(* IEC 61131-3 sources: daoli-st-library/DL_Device (part 34) *)

(* ---- FB_DL_VacuumEjector.st ---- *)
(*==============================================================================
 * 组件名称 (Component)  : FB_DL_VacuumEjector
 * 所属子库 (Sublibrary) : DL_Device
 * 当前版本 (Version)    : 1.0.1
 * 兼容性   (Platform)   : CODESYS 3.5 / TwinCAT 3 / 汇川 InoProShop / Machine Expert
 *                         仅依赖 Standard.library（TON / R_TRIG / TP），零厂商方言
 * 分类     (Category)   : 设备执行器功能块（Function Block，实现 I_DL_VacuumGenerator）
 * 功能简述 (Function)   : 真空发生器（射流式负压源）控制功能块。负压阈值
 *                         建立判据（负压域迟滞：建立用设定值、保持放宽
 *                         迟滞带防临界抖动）+ 可选真空开关双确认；破真空
 *                         吹气定宽单发脉冲（吹气期间真空阀强制断）；负压
 *                         反馈非有限值防御保持末次有效值；建立超时锁存；
 *                         状态机 ENUM + CASE + ELSE 兜底。
 * 接口实现 (Implements) : I_DL_VacuumGenerator。接口 OUT 列同名成员
 *                         （eState/bVacuumOk/fPressure/bFault/uErrorId）按
 *                         R22 以只读 PROPERTY GET 承载（内部镜像同源），
 *                         非接口成员 bVacuumValve/bBlowValve/bHolding 保留
 *                         VAR_OUTPUT；方法 CmdEvacuate/CmdBlowOff/CmdStop/
 *                         CmdReset 全部在本文件尾部落地。
 * 开源溯源 (Origin)     : 来源标签 lbp-device（RAW_NOTES_R6 S-1：真空吸持的
 *                         建立-保持迟滞判据、破真空吹气定宽脉冲、真空开关
 *                         双确认等行业公知工程惯例，公开教学资料，仅借鉴
 *                         通用工程语义；状态机、迟滞方向、故障码按本库红线
 *                         独立设计，clean-room 未复制源码）。
 * 红线自检 (Redline)    : R1 零全局变量表/外部变量引用 ✓｜R2 零物理 IO 地址 ✓
 *                         R3 纯 IEC 61131-3 ✓｜R4 防除零/非有限值防御/浮点
 *                         容差比较 ✓｜R5 全变量中英双语同行注释 ✓
 *                         R6 ENUM+CASE+ELSE ✓｜R7 六个定时器/边缘/脉冲实例
 *                         主体最前部无条件刷新 ✓
 * 公约遵循 (Convention) : 0.1/R23 本块为事件型状态机 + 逐拍组合阈值判定：
 *                         迟滞保持态每拍由实时负压重算自校正，无积分/滤波
 *                         类需要首扫初始化的连续量驻留状态，免首扫（无
 *                         bInit 标志）。
 *                         0.7 故障码段位 16#0003_xxxx：【故障级】0003_0230
 *                         负压反馈信号无效 / 0003_0231 真空建立超时（含
 *                         双确认模式下开关校验超窗）/ 0003_0232 非法状态，
 *                         全部 R15 锁存仅复位可清；本块无信息级码，bFault
 *                         派生式天然排除信息级（0.2）。
 * 偏离留档 (Deviation)  : 依 R11 头注释留档，共 1 条：
 *                         ① 规格建议吹气脉冲用"内部时间戳累积法"自实现
 *                           TP 语义；时间戳累积需时钟基准，与公约 0.9
 *                           "禁读时钟、时间一律注入"冲突，本实现改用
 *                           IEC 标准 TP 定宽脉冲定时器（Standard.library，
 *                           纯跨平台，语义等价），R14 断输入一拍规则对
 *                           组态期定值 PT 不涉及。
 * 修订历史 (Revision)   :
 *   2026-11-15  v1.0.0  首版入库（R6 轮 · DL_Device 阀门/驱动族深化）
 *   2026-11-15  v1.0.1  终审修复【致命】吹气脉冲触发时序：原实现 _bBlowReq
 *                       于主体末尾同拍自清，TP 实例（段 1 最前部刷新）永远
 *                       采不到 TRUE 入参，bBlowValve 恒 FALSE、eBlowing 态
 *                       下一拍即退回 eIdle（验收向量 V3 不成立，R13 逐拍
 *                       推演复现）。修法：自清动作移至 TP 实例调用之后，
 *                       TP 本拍采样 TRUE 起振、下一拍入参回落，定宽脉冲
 *                       由 TP 自身保持。引脚契约零变更。
 *============================================================================*)
FUNCTION_BLOCK FB_DL_VacuumEjector IMPLEMENTS I_DL_VacuumGenerator
VAR_INPUT
    bCmdEvacuate      : BOOL;           // 建立真空指令（Evacuate command），上升沿生效 / Evacuate command, rising edge effective
    bCmdBlowOff       : BOOL;           // 破真空吹气指令（Blow-off command），上升沿生效，输出 tBlowPulse 定宽脉冲 / Blow-off command, rising edge outputs fixed-width pulse
    fPressureFeedback : REAL;           // 负压表反馈（Pressure feedback）[kPa]，0=大气，负值=真空度；非有限值防御 / Pressure feedback [kPa], 0 = atmospheric, negative = vacuum, non-finite defended
    bFbVacuumSwitch   : BOOL;           // 可选真空开关反馈（Optional vacuum switch feedback），TRUE=真空确认 / Optional vacuum switch feedback, TRUE = vacuum confirmed
    bUseSensorCheck   : BOOL;           // 开关反馈校验使能（Sensor check enable），TRUE=负压阈值+开关双确认 / Sensor check enable, TRUE = threshold + switch dual confirmation
    fVacuumSetpoint   : REAL := -60.0;  // 真空建立阈值（Vacuum setpoint）[kPa]，负压域 / Vacuum establishment threshold in negative-pressure domain
    fVacuumHysteresis : REAL := 5.0;    // 真空判定迟滞（Vacuum hysteresis）[kPa]，保持判据放宽量，负值防御钳零 / Hysteresis band for hold criterion, negative clamped to zero
    tEstablishTimeout : TIME := T#5S;   // 真空建立超时（Establish timeout），T#0S=禁用 / Establish timeout, T#0S disables the check
    tBlowPulse        : TIME := T#500MS; // 破真空吹气脉冲宽度（Blow-off pulse width）/ Blow-off pulse width
    tDebounce         : TIME := T#20MS; // 开关反馈防抖（Switch debounce），T#0S=直通 / Switch feedback debounce, T#0S = pass-through
    bReset            : BOOL;           // 故障复位（Fault reset），上升沿生效 / Fault reset, rising edge effective
END_VAR

VAR_OUTPUT
    bVacuumValve : BOOL;                // 真空电磁阀输出（Vacuum solenoid valve），TRUE=抽真空 / Vacuum solenoid valve, TRUE = evacuating
    bBlowValve   : BOOL;                // 破真空吹气阀输出（Blow-off solenoid valve），定宽脉冲 / Blow-off solenoid valve, fixed-width pulse
    bHolding     : BOOL;                // 吸附保持中指示（Holding indicator），真空确认态为 TRUE / Holding indicator, TRUE in vacuum-ok state
END_VAR

VAR
    _eState         : E_DL_VacuumState := E_DL_VacuumState.eIdle; // 内部状态机步序（Internal state step），外部经属性只读 / Internal state, read-only via property
    _bFaultLatch    : BOOL;           // 故障锁存标志（Fault latch flag），仅复位清除 / Fault latch flag, cleared only by reset
    _uErrorIdInt    : UDINT;          // 内部故障码寄存（Internal error register），随锁存写入 / Internal error register written on latch
    _bPendEvac      : BOOL;           // 方法抽真空请求（Method evacuate request），由 CmdEvacuate 置位 / Method evacuate request set by CmdEvacuate
    _bPendBlow      : BOOL;           // 方法吹气请求（Method blow-off request），由 CmdBlowOff 置位 / Method blow-off request set by CmdBlowOff
    _bPendStop      : BOOL;           // 方法停止请求（Method stop request），由 CmdStop 置位 / Method stop request set by CmdStop
    _bPendReset     : BOOL;           // 方法复位请求（Method reset request），由 CmdReset 置位 / Method reset request set by CmdReset
    _bBlowReq       : BOOL;           // 吹气单拍触发请求（Blow pulse trigger request），上升沿消费置位一拍 / One-cycle blow trigger, set on edge consumption
    _fPressValid    : REAL := 0.0;    // 末次有效负压值（Last valid pressure）[kPa]，非有限值防御保持载体 / Last valid pressure hold carrier
    _fSetpEff       : REAL := -60.0;  // 防御后建立阈值（Sanitized setpoint）[kPa] / Sanitized vacuum setpoint
    _fHystEff       : REAL := 5.0;    // 防御后迟滞带（Sanitized hysteresis）[kPa]，钳制非负 / Sanitized hysteresis band, clamped non-negative
    _bPressValid    : BOOL;           // 本拍负压输入有效性（Pressure input validity this cycle），非有限值为 FALSE / FALSE when pressure input non-finite
    _bSwFilt        : BOOL;           // 防抖后真空开关（Debounced vacuum switch）/ Debounced vacuum switch signal
    _bInEstablish   : BOOL;           // 建立超时计时条件（Establish timeout timing condition）/ Timing condition of establish timeout
    _bEstToEn       : BOOL;           // 建立超时使能（Establish timeout enable），参数大于零有效 / Establish timeout enable, active when above zero
    _bEstablished   : BOOL;           // 本拍真空建立判据结果（Establishment criterion result this cycle）/ Establishment criterion result this cycle
    _bHoldCriterion : BOOL;           // 本拍保持判据结果（Hold criterion result this cycle），迟滞放宽域 / Hold criterion result within hysteresis band
    _fbTrigEvac     : R_TRIG;         // 引脚抽真空指令上升沿（Pin evacuate command edge）/ Pin evacuate command rising edge
    _fbTrigBlow     : R_TRIG;         // 引脚吹气指令上升沿（Pin blow-off command edge）/ Pin blow-off command rising edge
    _fbTrigReset    : R_TRIG;         // 引脚复位上升沿（Pin reset edge）/ Pin reset rising edge
    _fbTonSwDeb     : TON;            // 真空开关防抖定时器（Vacuum switch debounce timer）/ Vacuum switch debounce timer instance
    _fbTonEstablish : TON;            // 真空建立超时定时器（Establish timeout timer）/ Establish timeout timer instance
    _fbTpBlow       : TP;             // 吹气定宽脉冲定时器（Blow-off pulse timer），IEC 标准 TP / Blow-off fixed-width pulse timer, IEC standard TP
END_VAR

METHOD CmdEvacuate : BOOL
VAR_INPUT
END_VAR
IF _bFaultLatch OR (_eState = E_DL_VacuumState.eFault) THEN
    CmdEvacuate := FALSE;     // 故障态拒绝（Rejected in fault state）
ELSE
    _bPendEvac  := TRUE;      // 登记抽真空请求，主体状态机消化（Register evacuate request, consumed by body）
    CmdEvacuate := TRUE;      // 受理成功（Accepted）
END_IF

(*------------------------------------------------------------------------------
 * 方法: CmdBlowOff —— 破真空吹气指令（单发定宽脉冲）。故障态拒绝。
 *      Method CmdBlowOff - blow-off command (one-shot pulse), rejected in fault.
 *------------------------------------------------------------------------------*)
    END_METHOD

METHOD CmdBlowOff : BOOL
VAR_INPUT
END_VAR
IF _bFaultLatch OR (_eState = E_DL_VacuumState.eFault) THEN
    CmdBlowOff := FALSE;      // 故障态拒绝（Rejected in fault state）
ELSE
    _bPendBlow := TRUE;       // 登记吹气请求，主体状态机消化（Register blow request, consumed by body）
    CmdBlowOff := TRUE;       // 受理成功（Accepted）
END_IF

(*------------------------------------------------------------------------------
 * 方法: CmdStop —— 双阀全断保持现状。故障态拒绝返回 FALSE。
 *      Method CmdStop - both valves off and hold, rejected with FALSE in fault.
 *------------------------------------------------------------------------------*)
    END_METHOD

METHOD CmdStop : BOOL
VAR_INPUT
END_VAR
IF _bFaultLatch OR (_eState = E_DL_VacuumState.eFault) THEN
    CmdStop := FALSE;         // 故障态拒绝（Rejected in fault state）
ELSE
    _bPendEvac := FALSE;      // 注销全部动作请求（Cancel all action requests）
    _bPendBlow := FALSE;
    _bPendStop := TRUE;       // 登记停止请求，主体状态机消化（Register stop request, consumed by body）
    CmdStop    := TRUE;       // 受理成功（Accepted）
END_IF

(*------------------------------------------------------------------------------
 * 方法: CmdReset —— 复位故障，返回是否可复位（存在锁存故障时为 TRUE）。
 *      Method CmdReset - reset fault, returns TRUE only when a latch exists.
 *------------------------------------------------------------------------------*)
    END_METHOD

METHOD CmdReset : BOOL
VAR_INPUT
END_VAR
IF _bFaultLatch OR (_eState = E_DL_VacuumState.eFault) THEN
    _bPendReset := TRUE;      // 登记复位请求，主体状态机消化（Register reset request, consumed by body）
    CmdReset    := TRUE;      // 可复位（Resettable）
ELSE
    CmdReset    := FALSE;     // 无故障可复位（Nothing to reset）
END_IF

(*------------------------------------------------------------------------------
 * 属性: eState（GET）—— 当前状态机状态只读视图。
 *      Property eState (GET) - read-only view of the current state machine state.
 *------------------------------------------------------------------------------*)
    END_METHOD

// ============================================================================
// 段 1｜定时器与边缘检测实例无条件周期刷新（R7：严禁置于 IF/CASE 分支内）
//      Unconditional per-cycle refresh of all timer and edge instances (R7)
// ============================================================================
_fbTrigEvac(CLK := bCmdEvacuate);
_fbTrigBlow(CLK := bCmdBlowOff);
_fbTrigReset(CLK := bReset);
_fbTonSwDeb(IN := bFbVacuumSwitch, PT := tDebounce); // 开关持续为真 tDebounce 才确认（Switch must hold TRUE for tDebounce）
_bSwFilt := _fbTonSwDeb.Q;            // 防抖后开关（Debounced switch）
_bEstToEn := (tEstablishTimeout > T#0S); // 超时参数为零 = 自检禁用（Zero timeout = check disabled）
_bInEstablish := (_eState = E_DL_VacuumState.eEvacuating) AND _bEstToEn; // 建立超时计时条件（Timeout timing condition）
_fbTonEstablish(IN := _bInEstablish, PT := tEstablishTimeout);
_fbTpBlow(IN := _bBlowReq, PT := tBlowPulse); // 吹气定宽脉冲（Fixed-width blow pulse, TP semantics）
_bBlowReq := FALSE;                   // 单拍触发请求在 TP 采样后立即自清：TP 于本拍见到
                                      // TRUE 并起振，下一拍入参回落 FALSE，TP 定宽保持
                                      // （One-cycle trigger cleared right after TP sampling,
                                      // pulse held by TP for the full width）

// ============================================================================
// 段 2｜参数防御（0.8：非数自比检测，默认值先赋）+ 迟滞钳零
//      Parameter sanitation (0.8 NaN self-compare, defaults first) + clamp
// ============================================================================
_fSetpEff := fVacuumSetpoint;         // 建立阈值镜像（Setpoint mirror）
IF _fSetpEff <> _fSetpEff THEN        // 非数自比检测（NaN self-compare test）
    _fSetpEff := -60.0;               // 回落默认阈值（Fallback to default setpoint）
END_IF
_fHystEff := fVacuumHysteresis;       // 迟滞带镜像（Hysteresis mirror）
IF _fHystEff <> _fHystEff THEN        // 非数自比检测（NaN self-compare test）
    _fHystEff := 5.0;                 // 回落默认迟滞（Fallback to default hysteresis）
END_IF
IF _fHystEff < 0.0 THEN
    _fHystEff := 0.0;                 // 负迟滞会收窄判定域，钳零防错（Negative band narrows domain, clamp to zero）
END_IF

// ============================================================================
// 段 3｜负压输入有效性全局监视（优先级最高，吸附安全相关故为故障级）
//      Pressure validity global monitor (highest priority, fault level due
//      to holding safety relevance)
// ============================================================================
_bPressValid := (fPressureFeedback = fPressureFeedback); // 非数自比检测：等号成立即有效（NaN iff self-compare fails）
IF _bPressValid THEN
    _fPressValid := fPressureFeedback; // 更新末次有效负压（Update last valid pressure）
ELSE
    _bFaultLatch := TRUE;              // 反馈失效锁存（Feedback loss latch）
    _uErrorIdInt := 16#0003_0230;      // 0003_0230 负压反馈信号无效【故障级】/ Pressure feedback invalid, fault level
    _eState      := E_DL_VacuumState.eFault; // 强制故障态（Force fault state）
END_IF

// 真空判据（clean-room 内联迟滞语义，负压域方向：值越负真空越强）
// Vacuum criteria (inline hysteresis, negative-pressure domain: more negative = stronger)
_bEstablished := (_fPressValid <= _fSetpEff);                          // 建立判据：达到设定真空（Establish: reached setpoint vacuum）
_bHoldCriterion := (_fPressValid <= (_fSetpEff + _fHystEff));          // 保持判据：迟滞带放宽防临界抖动（Hold: widened by hysteresis band）

// ============================================================================
// 段 4｜核心状态机（ENUM + CASE，含 ELSE 非法状态兜底）
//      Core state machine (ENUM + CASE with ELSE illegal-state fallback)
// ============================================================================
IF _bFaultLatch OR (_eState = E_DL_VacuumState.eFault) THEN
    // 故障锁存态：清空全部请求，仅复位可退出（Latched fault: requests cleared, reset-only exit）
    _bPendEvac  := FALSE;             // 清方法请求（Clear method requests）
    _bPendBlow  := FALSE;
    _bPendStop  := FALSE;
    _bBlowReq   := FALSE;             // 撤销未触发脉冲请求（Cancel pending pulse trigger）
    IF _bPendReset OR _fbTrigReset.Q THEN
        _bPendReset  := FALSE;        // 消费复位请求（Consume reset request）
        _bFaultLatch := FALSE;        // 解除锁存（Release latch）
        _uErrorIdInt := 0;            // 故障码清零（Error code cleared）
        _eState      := E_DL_VacuumState.eIdle; // 回空闲态（Back to idle）
    END_IF
ELSE
    IF _bPendReset OR _fbTrigReset.Q THEN
        _bPendReset := FALSE;         // 无故障时消化复位请求（Absorb reset request when no fault）
    END_IF
    CASE _eState OF

        E_DL_VacuumState.eIdle: // 空闲稳态：双阀全断
            IF _bPendEvac OR _fbTrigEvac.Q THEN
                _bPendEvac := FALSE;            // 消费抽真空请求（Consume evacuate request）
                _eState    := E_DL_VacuumState.eEvacuating; // 转抽真空（To evacuating）
            ELSIF _bPendBlow OR _fbTrigBlow.Q THEN
                _bPendBlow := FALSE;            // 消费吹气请求（Consume blow request）
                _bBlowReq  := TRUE;             // 触发定宽脉冲（Trigger fixed-width pulse）
                _eState    := E_DL_VacuumState.eBlowing;
            ELSIF _bPendStop THEN
                _bPendStop := FALSE;            // 空闲态消化停止请求（Absorb stop request in idle）
            END_IF

        E_DL_VacuumState.eEvacuating: // 抽真空中：真空阀开，等待建立确认
            IF _bPendBlow OR _fbTrigBlow.Q THEN
                _bPendBlow := FALSE;            // 中途改吹气（Mid-way blow-off）
                _bBlowReq  := TRUE;
                _eState    := E_DL_VacuumState.eBlowing;
            ELSIF _bPendStop THEN
                _bPendStop := FALSE;            // 停止：双阀全断（Stop: both valves off）
                _eState    := E_DL_VacuumState.eIdle;
            ELSIF bUseSensorCheck AND _bEstablished AND (NOT _bSwFilt) THEN
                // 阈值达成但开关未确认：继续抽气等待（Threshold reached, switch pending: keep evacuating）
            ELSIF (NOT bUseSensorCheck) AND _bEstablished THEN
                _eState := E_DL_VacuumState.eVacuumOk; // 纯阈值模式：建立确认（Pure threshold: established）
            ELSIF bUseSensorCheck AND _bEstablished AND _bSwFilt THEN
                _eState := E_DL_VacuumState.eVacuumOk; // 双确认模式：阈值+开关齐备（Dual confirm: threshold AND switch）
            ELSIF _fbTonEstablish.Q THEN
                _bFaultLatch := TRUE;           // 建立超时锁存（Establish timeout latch）
                _uErrorIdInt := 16#0003_0231;   // 0003_0231 真空建立超时/反馈校验失败【故障级】/ Establish timeout or check failure, fault level
                _eState      := E_DL_VacuumState.eFault;
            END_IF

        E_DL_VacuumState.eVacuumOk: // 真空保持态：吸附保持中
            IF _bPendBlow OR _fbTrigBlow.Q THEN
                _bPendBlow := FALSE;            // 破真空放料（Release workpiece by blow-off）
                _bBlowReq  := TRUE;
                _eState    := E_DL_VacuumState.eBlowing;
            ELSIF _bPendStop THEN
                _bPendStop := FALSE;            // 停止：双阀全断（Stop: both valves off）
                _eState    := E_DL_VacuumState.eIdle;
            ELSIF NOT _bHoldCriterion THEN
                _eState := E_DL_VacuumState.eEvacuating; // 真空丢失（超迟滞带）：自动重建（Vacuum lost beyond band: auto re-establish）
            ELSIF bUseSensorCheck AND (NOT _bSwFilt) THEN
                _eState := E_DL_VacuumState.eEvacuating; // 双确认模式下开关脱开：自动重建（Switch dropped in dual mode: re-establish）
            END_IF

        E_DL_VacuumState.eBlowing: // 吹气中：吹气阀定宽脉冲，真空阀强制断
            IF _bPendBlow OR _fbTrigBlow.Q THEN
                _bPendBlow := FALSE;            // 吹气中重复触发忽略（Retrigger ignored while blowing）
            ELSIF _bPendStop THEN
                _bPendStop := FALSE;            // 停止请求提前截断脉冲（Stop request truncates pulse early）
                _bBlowReq  := FALSE;
                _eState    := E_DL_VacuumState.eIdle;
            ELSIF NOT _fbTpBlow.Q THEN
                _eState := E_DL_VacuumState.eIdle; // 脉冲宽度计满自动回空闲（Pulse completed, back to idle）
            END_IF

        ELSE // 非法状态兜底：任何越界枚举值强制锁存故障（Illegal state fallback）
            _bFaultLatch := TRUE;               // 故障锁存（Fault latched）
            _uErrorIdInt := 16#0003_0232;       // 0003_0232 非法状态【故障级】/ Illegal state, fault level
            _eState      := E_DL_VacuumState.eFault;
    END_CASE
END_IF

// ============================================================================
// 段 5｜阀输出推导 + 出口断言（硬约束：吹气期间真空阀必断；故障/空闲双阀必断）
//      Valve output derivation + exit assertions (vacuum valve forced off
//      while blowing; both valves off in fault/idle)
// ============================================================================
bVacuumValve := (_eState = E_DL_VacuumState.eEvacuating) OR (_eState = E_DL_VacuumState.eVacuumOk); // 抽真空与保持期真空阀开（Valve open while evacuating/holding）
bBlowValve := (_eState = E_DL_VacuumState.eBlowing) AND _fbTpBlow.Q; // 吹气阀随 TP 定宽脉冲（Blow valve follows TP pulse）
IF (_eState = E_DL_VacuumState.eBlowing) OR (_eState = E_DL_VacuumState.eFault)
   OR (_eState = E_DL_VacuumState.eIdle) THEN
    bVacuumValve := FALSE;              // 出口断言：吹气/故障/空闲真空阀必断（Assertion: vacuum valve off in blowing/fault/idle）
END_IF

(*------------------------------------------------------------------------------
 * 方法: CmdEvacuate —— 建立真空指令（单发）。故障态一律拒绝返回 FALSE。
 *      Method CmdEvacuate - evacuate command (one-shot), rejected with FALSE in fault.
 *------------------------------------------------------------------------------*)

PROPERTY eState : E_DL_VacuumState
eState := _eState;            // 返回内部状态（Return internal state）

(*------------------------------------------------------------------------------
 * 属性: bVacuumOk（GET）—— 真空建立确认（吸附保持态为 TRUE）。
 *      Property bVacuumOk (GET) - vacuum established (TRUE in holding state).
 *------------------------------------------------------------------------------*)
PROPERTY bVacuumOk : BOOL
bVacuumOk := (_eState = E_DL_VacuumState.eVacuumOk); // 显式状态派生式（Explicit state-derived form）

(*------------------------------------------------------------------------------
 * 属性: fPressure（GET）—— 负压反馈值 [kPa]，0=大气压，负值=真空度。
 *      Property fPressure (GET) - pressure feedback [kPa], 0 = atmospheric, negative = vacuum.
 *------------------------------------------------------------------------------*)
PROPERTY fPressure : REAL
fPressure := _fPressValid;    // 返回末次有效负压保持值（Return last valid pressure hold value）

(*------------------------------------------------------------------------------
 * 属性: bFault（GET）—— 故障锁存指示（信息级码不置本位，0.2 公约）。
 *      Property bFault (GET) - fault latch indicator, info-level codes excluded.
 *------------------------------------------------------------------------------*)
PROPERTY bFault : BOOL
bFault := _bFaultLatch OR (_eState = E_DL_VacuumState.eFault); // 显式排除信息级派生式（Explicit derived form excluding info codes）

(*------------------------------------------------------------------------------
 * 属性: uErrorId（GET）—— 末次故障码（0=无故障）。
 *      Property uErrorId (GET) - last error code (0 = none).
 *------------------------------------------------------------------------------*)
PROPERTY uErrorId : UDINT
uErrorId := _uErrorIdInt;     // 返回内部故障码寄存（Return internal error register）
END_FUNCTION_BLOCK

(* ---- FB_DL_VacuumPumpBasePress.st ---- *)
(*
  Component : FB_DL_VacuumPumpBasePress
  Category  : DL_Device
  Type      : FB
  Version   : 1.0.0
  CodeSeg   : 16#03_1_03
  Summary   : 真空泵本底压强与恢复时间台账：本底压强滑动平均平滑 + 起泵恢复超时事件计数留痕。
              Vacuum pump base pressure and recovery ledger: moving-average smoothing plus restart recovery timeout counting.
  溯源声明  : 道莅自研 clean-room
  边界安全  : 压强非物理域闸（负压 < 0 拦截，非有限 NaN/Inf 拦截）；MA 环形缓冲点数域闸（2..16，防越界）；
              采样窗/恢复窗时长正域闸（> 0）；MA 采样窗与恢复计时窗为独立 TON 实例；
              恢复超时计数用事件触发（timing 停止后不重复累加）；锁存故障有可达清码路径（恢复成功即清）。
  复用      : 无
*)

FUNCTION_BLOCK FB_DL_VacuumPumpBasePress
VAR_INPUT
    bRun       : BOOL;                  (* 监视使能 · Enable *)
    bPumpRun   : BOOL;                  (* 泵运行反馈 [开关]，上升沿起恢复计时 · Pump run feedback *)
    fPressKpa  : LREAL;                 (* 泵入口压强 [kPa] · Pump inlet pressure *)
    fBaseOkKpa : LREAL := 5.0;          (* 本底压强达标阈 [kPa] · Base pressure target *)
    tMaWinMs   : TIME  := T#2000MS;     (* MA 采样节拍 [ms] · MA sample pace *)
    tRecWinMs  : TIME  := T#60000MS;    (* 恢复计时窗 [ms] · Recovery timing window *)
    nMaPts     : INT   := 8;            (* MA 有效点数 [点]，域 2 到 16 · MA valid points *)
    fEps       : LREAL := 1.0E-6;       (* 浮点判零容差 [实数域] · Floating zero tolerance *)
END_VAR
VAR_OUTPUT
    fMaKpa      : LREAL;                (* 本底压强滑动平均 [kPa] · Moving average pressure *)
    bRecTiming  : BOOL;                 (* 恢复计时进行中 [开关] · Recovery timing active *)
    bRecOk      : BOOL;                 (* 最近一次恢复成功 [开关] · Last recovery succeeded *)
    nRecTimeout : UDINT;                (* 恢复超时累计 [次]，事件计数防回卷 · Recovery timeout count *)
    bError      : BOOL;                 (* 故障标志，与故障码配对 · Fault flag paired with codes *)
    uErrorId    : UDINT;                (* 事件码 16#0000_0103，0 无事件 · Event code *)
END_VAR
VAR
    uCode    : WORD;    (* 码位暂存，每拍重算 [码] · Code staging *)
    tonMa    : TON;     (* MA 采样节拍 [ms]，自复位振荡 · MA pace timer, self-reset *)
    tonRec   : TON;     (* 恢复计时窗 [ms]，独立实例 · Recovery window timer, separate instance *)
    rTrigRun : R_TRIG;  (* 起泵上升沿 · Pump start rising edge *)
    aRing    : ARRAY[1..16] OF LREAL;   (* MA 环形缓冲 [kPa] · MA ring buffer *)
    nHead    : INT;     (* 环形头下标 [索引] · Ring head index *)
    nFill    : INT;     (* 已填充点数 [点] · Filled point count *)
    fSum     : LREAL;   (* 环内累加和 [kPa] · Ring sum *)
    bRecFlt  : BOOL;    (* 恢复超时锁存 · Recovery timeout latched *)
    bSigOk   : BOOL;    (* 输入有效标志 · Input validity flag *)
    bTick    : BOOL;    (* 采样到点脉冲 [脉冲] · Sample tick pulse *)
    nI       : INT;     (* 求和循环下标 [索引] · Sum loop index *)
END_VAR
VAR CONSTANT
    DL_VBP_NMAX : INT := 16;            (* 环形缓冲容量 [点] · Ring capacity *)
END_VAR

(* === 段 0 · 实例刷新（每拍无条件，红线 7）=== *)
tonMa(IN := NOT tonMa.Q, PT := tMaWinMs);       (* 采样节拍自复位振荡 / Self-reset MA pace *)
tonRec(IN := bRecTiming, PT := tRecWinMs);      (* 恢复计时窗独立实例 / Separate recovery window *)
rTrigRun(CLK := bPumpRun);                      (* 起泵沿检测 / Pump start edge *)
bTick := tonMa.Q;                               (* 采样脉冲 / Sample tick *)

(* === 段 1 · 输入校验与量程闸 === *)
uCode := 16#0000;                       // 每拍清码（可达清零基线）/ Clear codes each scan
bSigOk := (fPressKpa = fPressKpa) AND (ABS(fPressKpa) < 1.0E308)    // 非有限拦截 / Non-finite guard
          AND (fPressKpa >= 0.0)                                     // 压强非负域闸 / Non-negative pressure
          AND (nMaPts >= 2) AND (nMaPts <= DL_VBP_NMAX)              // 点数域闸，防越界 / Point-count gate
          AND (tMaWinMs > T#0MS) AND (tRecWinMs > T#0MS);            // 窗时长正域闸 / Window duration gates
IF NOT bSigOk THEN
    uCode := 16#0103;                   // 故障级：域外，台账冻结 / Fault: domain invalid
END_IF

(* === 段 2 · 主逻辑：MA 平滑与恢复台账 === *)
IF bSigOk THEN
    IF bTick THEN                       (* 采样到点：写环并重算均值 / Sample tick: write ring *)
        IF nFill < nMaPts THEN
            nFill := nFill + 1;         (* 未满先增填充数 / Grow fill count *)
        ELSE
            fSum := fSum - aRing[nHead];    (* 满环先减旧值 / Remove the old value *)
        END_IF
        aRing[nHead] := fPressKpa;      (* 写入新采样 / Write the new sample *)
        fSum := fSum + fPressKpa;       (* 累加新值 / Add the new value *)
        nHead := (nHead MOD DL_VBP_NMAX) + 1;   (* 头下标循环推进 / Advance the head *)
    END_IF
    IF nFill >= 2 THEN
        fMaKpa := fSum / UDINT_TO_LREAL(INT_TO_UDINT(nFill));   (* 均值，填充数 ≥2 已闸 / Mean *)
    END_IF
    (* 恢复台账：起泵沿起计时，达标即成功，超窗即超时计数 / Recovery ledger *)
    IF rTrigRun.Q THEN
        bRecTiming := TRUE;             (* 拍 N 起泵沿进入，本拍置计时，拍 N+1 tonRec 生效 / Start timing *)
        bRecOk := FALSE;                (* 新恢复未达标 / New recovery pending *)
    END_IF
    IF bRecTiming AND (fMaKpa <= fBaseOkKpa) AND (nFill >= nMaPts) THEN
        bRecTiming := FALSE;            (* 达标：停止计时 / Reached target: stop timing *)
        bRecOk := TRUE;                 (* 恢复成功 / Recovery succeeded *)
        bRecFlt := FALSE;               (* 超时锁存清码（可达路径）/ Reachable clear of the latch *)
    END_IF
    IF bRecTiming AND tonRec.Q THEN     (* 计时窗满仍未达标 / Window expired without target *)
        bRecTiming := FALSE;            (* 停止计时，防重复计数 / Stop timing, no double count *)
        bRecFlt := TRUE;                (* 超时锁存 / Latch the timeout *)
        IF nRecTimeout < 4294967290 THEN
            nRecTimeout := nRecTimeout + 1;     (* 事件计数，一次恢复只计一次 / Count once per recovery *)
        END_IF
    END_IF
END_IF

(* === 段 3 · 输出映射与故障码 === *)
IF NOT bRun THEN
    bRecTiming := FALSE;                (* 撤使能停计时 / Stop timing on disable *)
END_IF
bError := bRecFlt OR (uCode <> 16#0000);        (* 故障标志：超时锁存或域外 / Fault flag *)
IF bRecFlt THEN
    uErrorId := WORD_TO_UDINT(16#0103); (* 码位 16#0000_0103 恢复超时锁存 / Recovery timeout code *)
ELSE
    uErrorId := WORD_TO_UDINT(uCode);   (* 域外码或零 / Domain code or zero *)
END_IF
END_FUNCTION_BLOCK

(* ---- FB_DL_ValveCycleCountBank.st ---- *)
//==============================================================================
// 功能块：FB_DL_ValveCycleCountBank ｜ 中文名称：多阀动作计数寿命台账组
// 所属子库：DL_Device ｜ 版本：v1.0.0 ｜ 日期：2026-11-23
// 兼容：CODESYS V3.5+ / TwinCAT 3 / 汇川 InoProShop（纯标准库 R_TRIG）
// 功能描述：4 阀动作计数寿命台账 Bank：每通道对阀指令上升沿计数（全行程
//           动作次数），独立维护阈值（UDINT），计数达阈值置该通道维护预警
//           bMaintX（不置故障——维护预警是台账事实非软件错误）。计数饱和
//           于 UDINT 上限 4294967295 不回绕（信息级留痕），复位经 bRst 沿
//           或 bRstChX 单通道沿。
//           同族分工：单阀寿命判定（阀位双阈值跨越 + 双源同证去抖 + 分级
//           预警）属 FB_DL_ValveCycleLifeCounter；本件为 4 通道指令沿计数
//           Bank 台账（无反馈口径），互不替代（R73 互引）。
// 开源溯源 (Origin)：原创实现（t2-2-lbp 阀诊断深化，零外部源码行，clean-room
//           独立编写）
// 公开接口清单：输入 {bCmdCh1..4, uLimitCh1..4} / bRst / bRstCh1..4；
//               输出 {uCntCh1..4, bMaintCh1..4} / uErrCode / bValid
// 错误码表：16#0003_0754 信息级（任一通道计数饱和不回绕，不置 bError）/
//           16#0003_0755 预留禁用（不得挪用）
// 状态机：N/A（台账计数无状态机；R_TRIG ×8 每拍无条件刷新）
// 边界行为：① 计数饱和于 4294967295 不回绕（信息级 0754 留痕）；
//           ② R_TRIG 全部每拍无条件刷新（不入分支，红线 R7）；
//           ③ 维护预警随计数回落自动撤销（阈值比较瞬时量，不锁存）；
//           ④ 复位沿仅清计数，不清阈值与信息码（信息码每拍重算）。
// 修订历史：v1.0.0 2026-11-23 首版（R73 派单 · 批 3 · 序 16）
//==============================================================================

(*==============================================================================
 * 功能块: FB_DL_ValveCycleCountBank
 * 调用约定: 每个扫描周期无条件调用一次；实例状态全部驻留于私有变量。
 *==============================================================================*)
FUNCTION_BLOCK FB_DL_ValveCycleCountBank
VAR_INPUT
    bCmdCh1  : BOOL := FALSE;          // 阀 1 指令（上升沿 = 一次全行程动作）/ Valve 1 command, rising edge = one full stroke
    bCmdCh2  : BOOL := FALSE;          // 阀 2 指令（上升沿计数）/ Valve 2 command, counted on rising edge
    bCmdCh3  : BOOL := FALSE;          // 阀 3 指令（上升沿计数）/ Valve 3 command, counted on rising edge
    bCmdCh4  : BOOL := FALSE;          // 阀 4 指令（上升沿计数）/ Valve 4 command, counted on rising edge
    uLimitCh1: UDINT := 1000000;       // 阀 1 维护阈值 [次] / Valve 1 maintenance threshold [cycles]
    uLimitCh2: UDINT := 1000000;       // 阀 2 维护阈值 [次] / Valve 2 maintenance threshold [cycles]
    uLimitCh3: UDINT := 1000000;       // 阀 3 维护阈值 [次] / Valve 3 maintenance threshold [cycles]
    uLimitCh4: UDINT := 1000000;       // 阀 4 维护阈值 [次] / Valve 4 maintenance threshold [cycles]
    bRst     : BOOL := FALSE;          // 全组复位（上升沿，清全部计数）/ Bank reset, rising edge, clears all counts
    bRstCh1  : BOOL := FALSE;          // 阀 1 单通道复位沿 / Valve 1 channel reset edge
    bRstCh2  : BOOL := FALSE;          // 阀 2 单通道复位沿 / Valve 2 channel reset edge
    bRstCh3  : BOOL := FALSE;          // 阀 3 单通道复位沿 / Valve 3 channel reset edge
    bRstCh4  : BOOL := FALSE;          // 阀 4 单通道复位沿 / Valve 4 channel reset edge
END_VAR
VAR_OUTPUT
    uCntCh1  : UDINT;                  // 阀 1 累计动作数 [次] / Valve 1 accumulated cycles
    uCntCh2  : UDINT;                  // 阀 2 累计动作数 [次] / Valve 2 accumulated cycles
    uCntCh3  : UDINT;                  // 阀 3 累计动作数 [次] / Valve 3 accumulated cycles
    uCntCh4  : UDINT;                  // 阀 4 累计动作数 [次] / Valve 4 accumulated cycles
    bMaintCh1: BOOL;                   // 阀 1 维护预警（计数达阈值）/ Valve 1 maintenance warning
    bMaintCh2: BOOL;                   // 阀 2 维护预警（计数达阈值）/ Valve 2 maintenance warning
    bMaintCh3: BOOL;                   // 阀 3 维护预警（计数达阈值）/ Valve 3 maintenance warning
    bMaintCh4: BOOL;                   // 阀 4 维护预警（计数达阈值）/ Valve 4 maintenance warning
    uErrCode : UDINT;                  // 信息级码，0 = 无信息 / Info-level code, 0 = none
    bValid   : BOOL;                   // 输出可用标志 / Outputs usable flag
END_VAR
VAR
    trigCmd1 : R_TRIG;                 // 阀 1 指令沿检测，每拍无条件刷新 / Valve 1 command edge, refreshed every scan
    trigCmd2 : R_TRIG;                 // 阀 2 指令沿检测，每拍无条件刷新 / Valve 2 command edge, refreshed every scan
    trigCmd3 : R_TRIG;                 // 阀 3 指令沿检测，每拍无条件刷新 / Valve 3 command edge, refreshed every scan
    trigCmd4 : R_TRIG;                 // 阀 4 指令沿检测，每拍无条件刷新 / Valve 4 command edge, refreshed every scan
    trigRst  : R_TRIG;                 // 全组复位沿检测，每拍无条件刷新 / Bank reset edge, refreshed every scan
    trigRst1 : R_TRIG;                 // 阀 1 复位沿检测，每拍无条件刷新 / Valve 1 reset edge, refreshed every scan
    trigRst2 : R_TRIG;                 // 阀 2 复位沿检测，每拍无条件刷新 / Valve 2 reset edge, refreshed every scan
    trigRst3 : R_TRIG;                 // 阀 3 复位沿检测，每拍无条件刷新 / Valve 3 reset edge, refreshed every scan
    trigRst4 : R_TRIG;                 // 阀 4 复位沿检测，每拍无条件刷新 / Valve 4 reset edge, refreshed every scan
END_VAR
VAR CONSTANT
    DL_VCC_MAX     : UDINT := 4294967295; // UDINT 计数上限（饱和不回绕）/ UDINT count ceiling, saturating
    DL_VCC_CODE_SAT: UDINT := 16#0003_0754; // 信息级：计数饱和码 / Info code: count saturated
END_VAR

// ---- 段 1｜沿实例无条件刷新（红线 R7：全部 8 实例不入分支）----
trigCmd1(CLK := bCmdCh1);             // 阀 1 指令沿每拍刷新 / Valve 1 edge refreshed
trigCmd2(CLK := bCmdCh2);             // 阀 2 指令沿每拍刷新 / Valve 2 edge refreshed
trigCmd3(CLK := bCmdCh3);             // 阀 3 指令沿每拍刷新 / Valve 3 edge refreshed
trigCmd4(CLK := bCmdCh4);             // 阀 4 指令沿每拍刷新 / Valve 4 edge refreshed
trigRst(CLK := bRst);                 // 全组复位沿每拍刷新 / Bank reset edge refreshed
trigRst1(CLK := bRstCh1);             // 阀 1 复位沿每拍刷新 / Valve 1 reset edge refreshed
trigRst2(CLK := bRstCh2);             // 阀 2 复位沿每拍刷新 / Valve 2 reset edge refreshed
trigRst3(CLK := bRstCh3);             // 阀 3 复位沿每拍刷新 / Valve 3 reset edge refreshed
trigRst4(CLK := bRstCh4);             // 阀 4 复位沿每拍刷新 / Valve 4 reset edge refreshed

// ---- 段 2｜计数推进：饱和不回绕（信息级留痕，每拍重算）----
IF trigCmd1.Q AND (uCntCh1 < DL_VCC_MAX) THEN
    uCntCh1 := uCntCh1 + 1;           // 阀 1 计数推进 / Valve 1 count advance
END_IF
IF trigCmd2.Q AND (uCntCh2 < DL_VCC_MAX) THEN
    uCntCh2 := uCntCh2 + 1;           // 阀 2 计数推进 / Valve 2 count advance
END_IF
IF trigCmd3.Q AND (uCntCh3 < DL_VCC_MAX) THEN
    uCntCh3 := uCntCh3 + 1;           // 阀 3 计数推进 / Valve 3 count advance
END_IF
IF trigCmd4.Q AND (uCntCh4 < DL_VCC_MAX) THEN
    uCntCh4 := uCntCh4 + 1;           // 阀 4 计数推进 / Valve 4 count advance
END_IF
IF (uCntCh1 = DL_VCC_MAX) OR (uCntCh2 = DL_VCC_MAX)
   OR (uCntCh3 = DL_VCC_MAX) OR (uCntCh4 = DL_VCC_MAX) THEN
    uErrCode := DL_VCC_CODE_SAT;      // 信息级：计数饱和不回绕留痕 / Info: saturation trace, no wrap
END_IF

// ---- 段 3｜复位路径：全组沿 + 单通道沿（锁存声明的清除沿）----
IF trigRst.Q THEN                     // 全组复位沿
    uCntCh1 := 0;                     // 阀 1 计数清零 / Valve 1 count cleared
    uCntCh2 := 0;                     // 阀 2 计数清零 / Valve 2 count cleared
    uCntCh3 := 0;                     // 阀 3 计数清零 / Valve 3 count cleared
    uCntCh4 := 0;                     // 阀 4 计数清零 / Valve 4 count cleared
END_IF
IF trigRst1.Q THEN
    uCntCh1 := 0;                     // 阀 1 单通道清零 / Valve 1 channel clear
END_IF
IF trigRst2.Q THEN
    uCntCh2 := 0;                     // 阀 2 单通道清零 / Valve 2 channel clear
END_IF
IF trigRst3.Q THEN
    uCntCh3 := 0;                     // 阀 3 单通道清零 / Valve 3 channel clear
END_IF
IF trigRst4.Q THEN
    uCntCh4 := 0;                     // 阀 4 单通道清零 / Valve 4 channel clear
END_IF

// ---- 段 4｜维护预警装配：阈值比较瞬时量（随计数回落自动撤销，不锁存）----
bMaintCh1 := uCntCh1 >= uLimitCh1;    // 阀 1 维护预警 / Valve 1 maintenance warning
bMaintCh2 := uCntCh2 >= uLimitCh2;    // 阀 2 维护预警 / Valve 2 maintenance warning
bMaintCh3 := uCntCh3 >= uLimitCh3;    // 阀 3 维护预警 / Valve 3 maintenance warning
bMaintCh4 := uCntCh4 >= uLimitCh4;    // 阀 4 维护预警 / Valve 4 maintenance warning
bValid := TRUE;                       // 台账输出恒可用 / Ledger outputs always usable
END_FUNCTION_BLOCK

(* ---- FB_DL_ValveCycleLifeCounter.st ---- *)
(*
  Name        : FB_DL_ValveCycleLifeCounter
  Category    : DL_Device
  Version     : 1.0.0
  Purpose     : 阀门动作循环寿命计数：行程到位 + 扭角峰值双源同证并经去抖确认才计一个循环，累计数达保养阈值即预警；/ Valve cycle-life counter: one cycle is counted only when both stroke-limit and torque sources agree and the agreement is debounce-confirmed; a maintenance warning is raised at the threshold
  溯源        : 借 t2-8-isa182·回路一致性 的分类/参数域组织，clean-room 实现
  Boundary    : ① 组态闸：保养阈值 < 1 / 去抖时间 <= 0 → 锁存故障（阈值 0 会使预警无意义）；
                ② 双源判据：行程与扭角须同拍同真（AND），单源漂移不会虚计（去抖再拦短时毛刺）；
                ③ 计数用净额单点写入 + 饱和上限（R28 防回绕），不使用 CTU 双向端；
                ④ 循环脉冲 _bCycC 内部置位 → 段 5 统一出口映射单拍（R187），CASE 内不直写出口；
                ⑤ 本件仅计数与预警，不执行保养联锁（属主边界）。
*)
TYPE E_DL_VclState :
(
    eIdle  := 0,                             (* 未使能 / Disabled *)
    eCount := 10,                            (* 寿命计数运行 / Counting *)
    eFault := 90                             (* 故障锁存相 / Fault latched *)
);
END_TYPE

TYPE E_DL_VclCause :
(
    eNone       := 0,                        (* 无故障成因 / No cause *)
    eCfgIllegal := 1,                        (* 组态非法：阈值/去抖越域 / Illegal config *)
    ePhaseBad   := 2                         (* 非法相位兜底 / Illegal phase fallback *)
);
END_TYPE

FUNCTION_BLOCK FB_DL_ValveCycleLifeCounter
VAR_INPUT
    bStrokeOk   : BOOL := FALSE;             (* 行程到位信号（限位开关/位控回读）[-] / Stroke limit reached *)
    bTorqueOk   : BOOL := FALSE;             (* 扭角峰值信号（扭矩/扭角判据回读）[-] / Torque-angle criterion met *)
    tDebounce   : TIME := T#200MS;           (* 双源同证去抖时长，域 > T#0S [ms] / Dual-source debounce time, > 0 *)
    nMaintLimit : UDINT := 100000;           (* 保养阈值（累计循环数），域 >= 1 [次] / Maintenance cycle threshold, >= 1 *)
    bEnable     : BOOL := TRUE;              (* 计数使能 [-] / Enable *)
    bReset      : BOOL := FALSE;             (* 复位命令，上升沿清计数与故障（保养完成侧清零亦可用）[-] / Reset command *)
END_VAR
VAR_OUTPUT
    nCycles     : UDINT;                     (* 累计动作循环数（净额，饱和）[次] / Accumulated cycles, saturated *)
    fCycPct     : REAL;                      (* 寿命消耗百分比 = 计数/阈值（饱和 0..100）[%] / Life consumed percentage *)
    bCycPulse   : BOOL;                      (* 本拍新增一个循环（单拍脉冲）[-] / One new cycle this scan *)
    bMaintWarn  : BOOL;                      (* 保养预警：累计数 >= 阈值（电平，复位沿清）[-] / Maintenance warning level *)
    eState      : E_DL_VclState;             (* 状态出口 / State outlet *)
    eCause      : E_DL_VclCause;             (* 故障成因出口（R190 归因唯一） / Fault cause outlet *)
    bError      : BOOL;                      (* 故障锁存标志 [-] / Fault latch flag *)
END_VAR
VAR
    _eState   : E_DL_VclState := E_DL_VclState.eIdle;    (* 内部相位（CASE 唯一写入目标） / Internal phase *)
    _eCause   : E_DL_VclCause := E_DL_VclCause.eNone;    (* 故障成因锁存量 / Latched cause *)
    rtReset   : R_TRIG;                      (* 复位沿实例，段 0 无条件调用 / Reset edge instance *)
    rtCyc     : R_TRIG;                      (* 去抖确认输出沿实例，段 0 无条件调用 / Debounced-cycle edge *)
    tonDeb    : TON;                         (* 双源同证去抖计时器（IN 由双源派生） / Dual-source debounce timer *)
    _bFault   : BOOL;                        (* 故障锁存位 / Latched fault bit *)
    _bCfgBad  : BOOL;                        (* 组态非法当拍量 / Illegal config this scan *)
    _bDual    : BOOL;                        (* 双源同证当拍量（行程 AND 扭角） / Dual-source agreement this scan *)
    _bCycC    : BOOL;                        (* 循环确认内部单拍量（出口统一映射，R187） / Cycle-confirmed internal pulse *)
END_VAR
VAR CONSTANT
    DL_VCL_EPS    : REAL  := 1.0E-6;         (* 判零容差 [-] / Epsilon *)
    DL_VCL_CNTMAX : UDINT := 4294967295;     (* 计数饱和上限（R28）[-] / Count saturation cap *)
    DL_VCL_PCTMAX : REAL  := 100.0;         (* 百分比满量程 [%] / Percentage full scale *)
END_VAR

(* —— 段 0：当拍判据派生 + 实例无条件刷新（R228A；R_TRIG/TON 全在段 0，无 IF 包裹） —— *)
_bCfgBad := (nMaintLimit < 1) OR NOT (tDebounce > T#0S);                       (* 阈值下限闸 + 去抖正域闸 / Threshold and debounce gates *)
rtReset(CLK := bReset);                                                        (* 复位沿每拍必调 / Reset edge every scan *)
rtCyc(CLK := tonDeb.Q);                                                        (* 去抖确认输出沿每拍必调 / Debounced edge every scan *)
_bDual := bStrokeOk AND bTorqueOk;                                             (* 双源同证：行程 AND 扭角（单源漂移不虚计） / Dual-source agreement *)
tonDeb(IN := (_eState = E_DL_VclState.eCount) AND _bDual, PT := tDebounce);    (* 去抖计时（eCount 相位闸：eIdle/eFault 不计时，上拍相位 1 拍延迟可接受） / Debounce with phase gate *)

(* —— 段 1：单拍量预清零（R107） —— *)
_bCycC := FALSE;                                                               (* 循环脉冲内部量预清 / Cycle pulse preset *)
bCycPulse := FALSE;                                                            (* 循环脉冲出口预清 / Cycle pulse outlet preset *)
bMaintWarn := FALSE;                                                           (* 预警位预清（仅计数分支按阈值置位） / Warn preset *)

(* —— 段 2：复位沿处理（作用域：清故障 + 清计数 + 清出口 + 迁 eIdle，R283 逐项声明） —— *)
IF rtReset.Q THEN
    _bFault := FALSE;                                                          (* 清故障锁存 / Clear fault *)
    _eCause := E_DL_VclCause.eNone;                                            (* 清成因 / Clear cause *)
    nCycles := 0;                                                              (* 清累计循环数出口 / Clear cycle count *)
    fCycPct := 0.0;                                                            (* 清寿命百分比出口 / Clear life percentage *)
    bMaintWarn := FALSE;                                                       (* 清保养预警出口 / Clear warn outlet *)
    _eState := E_DL_VclState.eIdle;                                            (* 迁未使能相 / Back to idle *)
END_IF

(* —— 段 3：组态故障锁存（锁存至复位沿，R189） —— *)
IF _bCfgBad AND NOT _bFault THEN
    _bFault := TRUE;                                                           (* 锁存故障位 / Latch fault *)
    _eCause := E_DL_VclCause.eCfgIllegal;                                      (* 成因：组态非法 / Cause: illegal config *)
    _eState := E_DL_VclState.eFault;                                           (* 同步迁故障相 / Migrate to fault *)
END_IF

(* —— 段 4：CASE 主状态机（ELSE 兜底迁 eFault，红线 6） —— *)
CASE _eState OF
    E_DL_VclState.eIdle:                                                       (* 未使能：不计数，出口保持 0 语义 / Disabled *)
        nCycles := 0;                                                          (* 失能清计数出口（防隐性回夹） / Clear count outlet *)
        fCycPct := 0.0;                                                        (* 失能清百分比出口 / Clear percentage outlet *)
        bMaintWarn := FALSE;                                                   (* 失能清预警出口 / Clear warn outlet *)
        IF bEnable AND NOT _bFault THEN
            _eState := E_DL_VclState.eCount;                                   (* 使能进入计数 / Enter counting *)
        END_IF
    E_DL_VclState.eCount:                                                      (* 计数相：去抖确认后入账 / Counting *)
        IF NOT bEnable THEN
            _eState := E_DL_VclState.eIdle;                                    (* 失能回未使能 / Back to idle *)
        END_IF
        IF rtCyc.Q THEN                                                        (* 双源同证保持满去抖时长：确认一个循环 / Debounce elapsed: one cycle confirmed *)
            _bCycC := TRUE;                                                    (* 循环脉冲内部置位（出口统一映射，R187） / Cycle pulse internal *)
            IF nCycles < DL_VCL_CNTMAX THEN
                nCycles := nCycles + 1;                                        (* 计数净额 +1（饱和防回绕，R28） / Net +1, saturated *)
            END_IF
            IF nCycles >= nMaintLimit THEN
                bMaintWarn := TRUE;                                            (* 累计数达保养阈值：预警锁存（复位沿清） / Maintenance threshold reached *)
            END_IF
            fCycPct := UDINT_TO_REAL(nCycles) / UDINT_TO_REAL(nMaintLimit) * DL_VCL_PCTMAX;   (* 寿命消耗比：除子阈值 >= 1 由组态闸保证 [%] / Life ratio, divisor gated *)
            IF fCycPct > DL_VCL_PCTMAX THEN
                fCycPct := DL_VCL_PCTMAX;                                      (* 百分比上限饱和（该变量最后一次写，钳位不被覆盖） / Upper saturation, last write *)
            END_IF
        END_IF
        IF bMaintWarn = FALSE THEN
            IF nCycles >= nMaintLimit THEN                                     (* 达阈值后维持预警电平（阈值随组态下调亦能覆盖） / Hold warn level *)
                bMaintWarn := TRUE;                                            (* 预警电平保持 / Warn level held *)
            END_IF
        END_IF
    E_DL_VclState.eFault:                                                      (* 故障相：冻结保持末值，仅复位沿出 / Fault *)
        ;                                                                      (* 锁存回放（R28） / Replay from latch *)
    ELSE                                                                       (* 非法相位兜底迁安全态 / Illegal phase fallback *)
        _eState := E_DL_VclState.eFault;                                       (* 迁故障相 / To fault *)
        _bFault := TRUE;                                                       (* 同步锁存 / Latch *)
        _eCause := E_DL_VclCause.ePhaseBad;                                    (* 成因：非法相位 / Cause: illegal phase *)
END_CASE

(* —— 段 5：出口映射（内部 _b* → 输出单拍，R187；名实双出口，R191） —— *)
bCycPulse := _bCycC;                                                           (* 循环脉冲单拍出口 / Cycle pulse single-scan outlet *)
bError := _bFault;                                                             (* 故障标志镜像 / Fault flag mirror *)
eState := _eState;                                                             (* 状态出口 / State outlet *)
eCause := _eCause;                                                             (* 成因出口 / Cause outlet *)
END_FUNCTION_BLOCK

(* ---- FB_DL_ValveIslandDiag.st ---- *)
(*==============================================================================
 * 组件名称 (Component)  : FB_DL_ValveIslandDiag
 * 所属子库 (Sublibrary) : DL_Device
 * 当前版本 (Version)    : 1.0.0
 * 兼容性   (Platform)   : CODESYS 3.5 / TwinCAT 3 / 汇川 InoProShop / Machine Expert
 *                         仅依赖 Standard.library（TON / R_TRIG），零厂商方言
 * 来源标签 (Source)     : self-std（设备族新增线）
 * 功能描述 (Function)   : 阀岛（多阀槽位集束）诊断：①槽位占用仲裁——配置占用槽数与
 *                         实际上线槽数比对；②公共供气压力监视（欠压确认延时）；
 *                         ③逐槽位失联分类码位图与失联计数。
 * 分工互引 (Boundary)   : 单阀体机械 / 电气故障归 FB_DL_ControlValveDiag 与
 *                         FB_DL_PneuCylinderDiag；本件只做**阀岛级公共资源与槽位
 *                         上线状态**诊断，不下沉到单阀动作判定。
 * 边界与语义披露 (Boundary disclosure) :
 *   1) 槽位定长 8（DL_VI_SLOTS），越界无路径：nSlotUsed 域 1..8 由组态闸挡住，
 *      位图输出 uLostMask 的 bit i 对应槽位 i（bit0 = 槽位 0）。
 *   2) 占用仲裁口径：nSlotUsed 为组态占用数，实际上线数为 abSlotCommOk 为真的槽位数；
 *      上线数少于占用数即判失联（差值即 uLostMask 的置位数），多出的「超出占用」
 *      槽位为信息级占用冲突（不是故障，可能是有意扩展）。
 *   3) 公共供气压力欠压与槽位失联各自独立确认窗与独立码位（R190 归因唯一）；
 *      失联计数 nSlotsLost 为饱和计数（上限 8，结构上不会越界）。
 *   4) 非有限压力信号不参与欠压判据（保持上一拍确认状态），由信号闸置信息码，
 *      不锁存、不因一扫 NaN 让诊断永久失效。
 * 故障码表 (Error codes) :
 *   16#0003_0536 [故障级] 组态非法（占用槽数越域 / 压力阈 / 两确认窗）
 *                 反证：诊断挂起与「全部槽位正常且压力正常」输出组合相同。
 *   16#0003_0537 [故障级] 公共供气压力欠压确认，锁存至复位沿 + 压力恢复
 *                 反证：欠压与单槽失联都表现为「阀岛不可用」，处置不同（气源 vs 通讯）。
 *   16#0003_0538 [故障级] 槽位失联确认（上线数少于占用数），锁存至复位沿 + 恢复
 *                 反证：失联位图每拍刷新会掩盖「曾经失联」事实，锁存是唯一历史出口。
 *   16#0003_0483 [信息级] 上线槽位数多于配置占用数（占用冲突，按扩展容忍）
 *                 反证：多槽上线与「恰好全部占用上线」的输出差异只在配置侧，
 *                 运行期输出组合相同，无码不可观测。
 * 码位总账 (Code ledger) : 16#0003_0536 / 0537 / 0538 用 ｜ 16#0003_0483 用
 * 依赖     (Depends)    : 无 DL_ 内部依赖；Standard.library: TON / R_TRIG
 * 红线自检 (Redline)    : R1 ✓ 零全局变量 ｜ R2 ✓ 零 %I/%Q ｜ R3 ✓ 纯 IEC 61131-3
 *                         R4 ✓ 数组定长无越界 / 非有限三判 / 域闸全枚举
 *                         R5 ✓ 全变量双语同行注释 ｜ R6 ✓ 四态 ENUM + ELSE 兜底
 *                         R7 ✓ 一沿四计时主体最前部无条件刷新
 * 修订历史 (Revision)   : 2026-11-22  v1.0.0  首版入库（R69 构建轮 · 批 2 · N5）
 *============================================================================*)

(*-----------------------------------------------------------------------------
 * 枚举: E_DL_ValveIslandState（归属 DL_Device，与 FB_DL_ValveIslandDiag 同文件）
 *----------------------------------------------------------------------------*)
TYPE E_DL_ValveIslandState :
(
    eIdle    := 0,    // 未使能：诊断挂起 / Disabled, diagnosis suspended
    eWatch   := 10,   // 监视中：压力与槽位确认计时 / Watching, pressure and slot timers
    eAlarm   := 20,   // 已确认异常（至少一项锁存）/ Alarm latched
    eFault   := 99    // 组态非法：诊断拒绝 / Config illegal, diagnosis refused
);
END_TYPE

(*==============================================================================
 * 功能块: FB_DL_ValveIslandDiag
 * 调用约定: 每个扫描周期无条件调用一次。
 *============================================================================*)
FUNCTION_BLOCK FB_DL_ValveIslandDiag
VAR_INPUT
    abSlotCommOk  : ARRAY[0..7] OF BOOL;   // 逐槽位上线（通讯 OK）：bit i 对应槽位 i / per-slot online flags
    nSlotUsed     : INT := 8;              // 组态占用槽位数 [个]，域 1..8 / configured occupied slots, 1 to 8
    fSupplyPress  : REAL;                  // 公共供气压力 [bar] / common supply pressure [bar]
    fPressMin     : REAL := 4.0;           // 供气压力下限 [bar]，<= 0 组态非法 / supply pressure floor [bar]
    tPressConfirm : TIME := T#3S;          // 欠压确认窗 [s] / low-pressure confirm window [s]
    tSlotConfirm  : TIME := T#5S;          // 槽位失联确认窗 [s] / slot-loss confirm window [s]
    bEnable       : BOOL := TRUE;          // 使能 / enable
    bReset        : BOOL;                  // 上升沿：清欠压 / 失联锁存 / rising edge clears the latches
END_VAR
VAR_OUTPUT
    uLostMask     : WORD;                  // 逐槽失联位图（bit i = 槽位 i）/ per-slot loss bitmap
    nSlotsLost    : INT;                   // 失联槽位数 [个]，0..8 / lost slot count
    bSlotLost     : BOOL;                  // 槽位失联锁存（确认后常驻）/ slot loss latched
    bPressLow     : BOOL;                  // 供气欠压锁存 / low supply pressure latched
    bError        : BOOL;                  // 故障标志（组态 / 两类锁存归并）/ fault flag
    uErrorId      : UDINT;                 // 故障码，0 = 无故障 / error code, 0 = none
    eState        : E_DL_ValveIslandState; // 当前状态（供 HMI 诊断）/ current state
END_VAR
VAR
    fbTrigReset   : R_TRIG;                // 复位沿检测实例 / reset edge detector
    tonPress      : TON;                   // 欠压确认计时实例 / low-pressure confirm timer
    tonSlot       : TON;                   // 槽位失联确认计时实例 / slot-loss confirm timer
    eStateInt     : E_DL_ValveIslandState; // 主状态机内部当前态 / internal state
    nOnlineCnt    : INT;                   // 本拍上线槽位数 [个] / online slot count this scan
    nIdx          : INT;                   // 槽位遍历游标 [槽号] / slot cursor
    uMaskInt      : WORD;                  // 本拍失联位图累加 / loss bitmap accumulator
    bSlotCond     : BOOL;                  // 本拍失联判据成立 / slot-loss criterion true
    bPressCond    : BOOL;                  // 本拍欠压判据成立 / low-pressure criterion true
    bPressBad     : BOOL;                  // 压力信号非有限 / pressure non-finite
    bSlotLatch    : BOOL;                  // 失联锁存内部副本 / internal slot-loss latch
    bPressLatch   : BOOL;                  // 欠压锁存内部副本 / internal low-pressure latch
    bCfgBad       : BOOL;                  // 本拍组态非法 / config illegal this scan
    bCfgLatch     : BOOL;                  // 组态锁存（复位沿 + 组态改对解除）/ config latch
    bErrorInt     : BOOL;                  // 本拍故障置位累加 / fault set accumulator
    bFirstScan    : BOOL := TRUE;          // 上电首扫标志 / first-scan flag
END_VAR
VAR CONSTANT
    DL_VI_SLOTS   : INT := 8;              // 槽位定长 [个]，与数组维度一致 / fixed slot count
    DL_VI_FIN_LIM : REAL := 1.0E30;        // REAL 幅值兜底判界 / REAL magnitude bound
    DL_VI_BIT1    : WORD := 1;             // 位图基元（bit0 掩码）/ bitmap base element
END_VAR

(*------------------------------------------------------------------------------
 * 段 1｜无条件刷新区（红线 R7）：一沿二计时位于主体最前部
 *      Unconditional refresh: one edge and two timers at the very top
 *-----------------------------------------------------------------------------*)
fbTrigReset(CLK := bReset);

(* 段 2｜每拍预清（FB32-1）：单拍标志与位图累加量 / per-scan preset *)
bErrorInt := FALSE;
uMaskInt  := 16#0000;              // 失联位图每拍重算（事实量，非锁存）/ loss bitmap recomputed each scan
nOnlineCnt := 0;

(* 段 3｜上电首扫：锁存与状态落安全侧 / first-scan init *)
IF bFirstScan THEN
    eStateInt  := E_DL_ValveIslandState.eIdle;
    bSlotLatch := FALSE;
    bPressLatch := FALSE;
    bFirstScan := FALSE;
END_IF

(*------------------------------------------------------------------------------
 * 段 4｜组态域闸（R151 全枚举）+ 解除路径（R152 自证可达）
 *      Config gate plus the provably reachable clear path
 *-----------------------------------------------------------------------------*)
bCfgBad := (nSlotUsed < 1) OR (nSlotUsed > DL_VI_SLOTS)
           OR (fPressMin <= 0.0) OR (fPressMin <> fPressMin)
           OR (tPressConfirm <= T#0S) OR (tSlotConfirm <= T#0S);
IF bCfgBad THEN
    bCfgLatch := TRUE;
END_IF
IF fbTrigReset.Q AND (NOT bCfgBad) THEN
    bCfgLatch := FALSE;              // 组态锁存解除 / config latch cleared
    uErrorId  := 16#0000_0000;       // 码位随解除归零 / code cleared with the latch
END_IF
IF bCfgLatch THEN
    uErrorId  := 16#0003_0536;       // 故障级：组态非法 / fault: illegal configuration
    bErrorInt := TRUE;               // R45 配对 / paired with the code
    eStateInt := E_DL_ValveIslandState.eFault;
END_IF

(*------------------------------------------------------------------------------
 * 段 5｜占用仲裁：逐槽位统计上线数并构造失联位图（定长 FOR，无越界路径）
 *      Occupation arbitration: count online slots and build the loss bitmap
 *-----------------------------------------------------------------------------*)
FOR nIdx := 0 TO (DL_VI_SLOTS - 1) DO
    IF abSlotCommOk[nIdx] THEN
        nOnlineCnt := nOnlineCnt + 1;                        // 上线计数推进 [个] / online count up
    ELSIF nIdx < nSlotUsed THEN
        uMaskInt := uMaskInt OR SHL(DL_VI_BIT1, nIdx);       // 占用槽且离线：置失联位（nIdx <= 7 < 16 位宽，R48 归一）/ set the loss bit
    END_IF
END_FOR

bSlotCond  := nOnlineCnt < nSlotUsed;              // 上线数少于占用数即失联 / fewer online than occupied
bPressBad  := (fSupplyPress <> fSupplyPress)
              OR ((fSupplyPress - fSupplyPress) <> (fSupplyPress - fSupplyPress))
              OR (ABS(fSupplyPress) >= DL_VI_FIN_LIM);
bPressCond := (NOT bPressBad) AND (NOT bCfgLatch) AND (fSupplyPress < fPressMin);

IF (NOT bPressBad) AND (nOnlineCnt > nSlotUsed) THEN
    uErrorId := 16#0003_0483;      // 信息级：超出占用的槽位已上线（按扩展容忍）/ info: extra slots online
END_IF

(* 确认计时器门控：判据 AND 未锁存 AND 非组态故障（R99） *)
tonPress(IN := bPressCond AND (NOT bPressLatch), PT := tPressConfirm);
tonSlot(IN := bSlotCond AND (NOT bSlotLatch) AND (NOT bCfgLatch), PT := tSlotConfirm);

(*------------------------------------------------------------------------------
 * 段 6｜主状态机（红线 R6）：ENUM + CASE + ELSE 兜底
 *-----------------------------------------------------------------------------*)
CASE eStateInt OF

    E_DL_ValveIslandState.eIdle:
        IF bEnable AND (NOT bCfgLatch) THEN
            eStateInt := E_DL_ValveIslandState.eWatch;
        END_IF

    E_DL_ValveIslandState.eWatch:
        IF (NOT bEnable) OR bCfgLatch THEN
            eStateInt := E_DL_ValveIslandState.eIdle;
        ELSIF bSlotLatch OR bPressLatch THEN
            eStateInt := E_DL_ValveIslandState.eAlarm;       // 任一确认即告警驻留 / any confirmation alarms
        END_IF

    E_DL_ValveIslandState.eAlarm:
        (* 解除路径（R152 自证可达）：复位沿 AND 两判据本拍均已消失 AND 组态合法 *)
        IF fbTrigReset.Q AND (NOT bSlotCond) AND (NOT bPressCond) AND (NOT bCfgBad) THEN
            bSlotLatch  := FALSE;                            // 两类锁存同沿解除 / both latches cleared
            bPressLatch := FALSE;
            uErrorId    := 16#0000_0000;
            eStateInt   := E_DL_ValveIslandState.eWatch;
        ELSIF (NOT bEnable) OR bCfgLatch THEN
            eStateInt   := E_DL_ValveIslandState.eIdle;
        END_IF

    E_DL_ValveIslandState.eFault:
        IF fbTrigReset.Q AND (NOT bCfgBad) THEN
            bCfgLatch := FALSE;
            uErrorId  := 16#0000_0000;
            eStateInt := E_DL_ValveIslandState.eIdle;
        END_IF

    ELSE
        (* 非法状态拦截 / illegal state interception *)
        eStateInt := E_DL_ValveIslandState.eFault;
        uErrorId  := 16#0003_0536;
        bErrorInt := TRUE;

END_CASE;

(*------------------------------------------------------------------------------
 * 段 7｜确认到期消化：两类各自独立锁存 + 独立码位（R190 归因唯一）
 *      Confirm expiry digestion with two distinct codes
 *-----------------------------------------------------------------------------*)
IF tonPress.Q AND (NOT bPressLatch) THEN
    bPressLatch := TRUE;             // 欠压锁存 / low pressure latched
    uErrorId    := 16#0003_0537;     // 故障级：供气欠压确认 / fault: low supply pressure confirmed
    bErrorInt   := TRUE;             // R45 配对 / paired with the code
    eStateInt   := E_DL_ValveIslandState.eAlarm;
END_IF
IF tonSlot.Q AND (NOT bSlotLatch) THEN
    bSlotLatch := TRUE;              // 失联锁存 / slot loss latched
    uErrorId   := 16#0003_0538;      // 故障级：槽位失联确认 / fault: slot loss confirmed
    bErrorInt  := TRUE;              // R45 配对 / paired with the code
    eStateInt  := E_DL_ValveIslandState.eAlarm;
END_IF

(*------------------------------------------------------------------------------
 * 段 8｜输出单一出口（范式 P-05）
 *      Single output exit
 *-----------------------------------------------------------------------------*)
uLostMask  := uMaskInt;              // 失联位图直出（bit i = 槽位 i）/ loss bitmap straight out
(* 失联数 = 占用数 − 上线数（负值钳 0，结构上 nOnlineCnt <= 8 已由定长循环封顶）*)
(* Lost count equals occupied minus online, floored at zero *)
IF nOnlineCnt < nSlotUsed THEN
    nSlotsLost := nSlotUsed - nOnlineCnt;   // 失联槽位数 [个] / lost slot count
ELSE
    nSlotsLost := 0;                        // 无失联 [个] / no lost slot
END_IF
bSlotLost  := bSlotLatch;
bPressLow  := bPressLatch;
bError     := bErrorInt OR bCfgLatch OR (eStateInt = E_DL_ValveIslandState.eAlarm);
eState     := eStateInt;
END_FUNCTION_BLOCK

(* ---- FB_DL_ValvePartialStrokeTest.st ---- *)
(*
  组件名 Component   : FB_DL_ValvePartialStrokeTest
  子库 Sublibrary    : DL_Device
  版本 Version       : 1.0.0
  兼容性 Platform    : CODESYS 3.5 / TwinCAT 3 / 汇川 InoProShop / Machine Expert（仅 Standard.library）
  功能 Function      : 安全阀部分行程测试 PST 顺控：
                       1) 测试许可联锁：bProcessPermissive 为测试前置硬闸，许可撤销
                       即中止测试并锁存（过程条件优先于测试）；
                       2) 测试行程限幅：测试目标位钳制在 [fTestLoPct, fTestHiPct]
                       测试带内，钳位后照常执行（行程受限是 PST 的安全本意）；
                       3) 顺控：eIdle → eCheck（许可与组态闸）→ eMove（开阀到测试
                       目标位）→ eReturn（回正常位）→ eDone，各相超时独立 TON；
                       4) 测试结果判级：行程到位差 <= fTravelTolPct → 合格；短行程
                       超容差 → 降级（NE107 需要维护）；完全不动 → 失效。
                       NE107 健康出口引用唯一属主 E_DL_Ne107Status（零重声明）。
  边界 Boundary      : ① 本件只出阀位指令与健康等级，不写物理 IO；
                       ② NE107 枚举全库唯一属主在 DL_Device（DeviceHealthArbiter 文件），
                       本件只引用；eFailure 与故障锁存配对，bReset 上升沿解除；
                       ③ 故障锁存解除唯一路径 = bReset 上升沿（输入引脚，恒可达）；
                       ④ 无全局变量引用、无外部变量声明、无物理地址寻址。
  依赖 Depends       : E_DL_Ne107Status（DL_Device 唯一属主）；Standard.library（R_TRIG / TON）
  溯源 Origin        : 道莅自研 clean-room（参考 t2-8-ne107/ISA PST 语义分类与参数域，
                       零代码行复制；健康出口仅引用唯一属主枚举）
  码位 Code          : 16#03_2_F（Device 05xx 副带 052F）
  码表 Error codes（Device 故障窗口 052F，本件无信息码，单故障总码 + 成因枚举归因）:
    16#0003_052F 故障级：PST 故障总码（许可撤销 / 目标位超时 / 回位超时 /
                 组态非法 / 输入非有限），锁存至 bReset 上升沿，归因见 eCause
  修订历史 Revision  :
    2026-11-19  v1.0.0  R44 首版（批次 3 · 序号 11）
*)

TYPE E_DL_PstState :
(
    eIdle   := 0,   // 空闲：等测试沿 / Idle, waiting test edge
    eCheck  := 10,  // 检查：许可与组态闸 / Checking permissive and configuration
    eMove   := 20,  // 行程：开阀至测试目标位 / Moving to test target position
    eReturn := 30,  // 回程：回正常位 / Returning to normal position
    eDone   := 40,  // 完成：判级驻留 / Done, grading held
    eFault  := 90   // 故障：PST 锁存 / Fault, latched
);
END_TYPE

TYPE E_DL_PstCause :
(
    eNone       := 0,  // 无故障成因 / No cause
    ePermissive := 1,  // 测试许可撤销 / Test permissive lost
    eMoveTo     := 2,  // 目标位超时未到位 / Move target timeout
    eReturnTo   := 3,  // 回位超时未到位 / Return timeout
    eCfgIllegal := 4,  // 组态非法 / Illegal configuration
    eNonFinite  := 5   // 输入非有限 / Non-finite input
);
END_TYPE

FUNCTION_BLOCK FB_DL_ValvePartialStrokeTest
VAR_INPUT
    bEnable        : BOOL;               // 使能（电平）[-] / Enable
    bReset         : BOOL;               // 上升沿清故障锁存 [-] / Reset edge
    bTestCmd       : BOOL;               // 测试指令（上升沿承载）[-] / Test command edge
    bProcessPermissive: BOOL;            // 过程测试许可（硬联锁）[-] / Process test permissive
    fActPosPct     : REAL;               // 阀实际位置 [%] / Valve actual position
    fTestTargetPct : REAL;               // 测试目标位（会被钳入测试带）[%] / Test target position
    fNormalPosPct  : REAL := 0.0;        // 正常工作位 [%] / Normal operating position
    fTestLoPct     : REAL := 10.0;       // 测试带下限 [%] / Test band floor
    fTestHiPct     : REAL := 30.0;       // 测试带上限 [%] / Test band ceiling
    fTravelTolPct  : REAL := 2.0;        // 行程到位容差 [%] / Travel tolerance
    tMoveTo        : TIME := T#30S;      // 行程超时 [毫秒] / Move timeout
    tReturnTo      : TIME := T#30S;      // 回程超时 [毫秒] / Return timeout
END_VAR
VAR_OUTPUT
    fValveCmdPct   : REAL;               // 阀位指令输出 [%] / Valve position command
    bTestActive    : BOOL;               // 测试进行中电平 [-] / Test active level
    bTestPass      : BOOL;               // 结论：合格 [-] / Verdict pass flag
    bTestDerated   : BOOL;               // 结论：降级（短行程）[-] / Verdict derated flag
    fTestTravelPct : REAL;               // 实测测试行程 [%] / Measured test travel
    eNe107         : E_DL_Ne107Status;   // NE107 健康出口（唯一属主枚举） / NE107 health outlet
    eState         : E_DL_PstState;      // 状态出口，段尾单点映射 / State outlet
    eCause         : E_DL_PstCause;      // 故障成因出口（R190） / Fault cause outlet
    bError         : BOOL;               // 故障锁存标志 [-] / Fault latch flag
    uErrId         : UDINT;              // 事件码，0 = 无事件 / Event code
END_VAR
VAR
    rtReset: R_TRIG;                     // 复位沿实例，段 0 无条件刷新 / Reset edge
    rtTest : R_TRIG;                     // 测试沿实例，段 0 无条件刷新 / Test edge
    tonMoveTo : TON;                     // 行程超时（专用超时件命名） / Move timeout
    tonReturnTo: TON;                    // 回程超时（专用超时件命名） / Return timeout
    _eState: E_DL_PstState := E_DL_PstState.eIdle;     // 内部相位（CASE 唯一写入目标）/ Internal phase
    _eCause: E_DL_PstCause := E_DL_PstCause.eNone;     // 故障成因锁存（锁存量）/ Latched cause
    _fTargetUse: REAL;                   // 钳位后测试目标位 [%] / Clamped test target
    _fPosStart : REAL;                   // 测试起点位置 [%] / Test start position
    _bFault: BOOL;                       // 故障锁存位（锁存量） / Latched fault bit
    _uFault: UDINT;                      // 故障码锁存（锁存量） / Latched fault code
    _bCfgBad: BOOL;                      // 组态非法当拍量 [-] / Config illegal flag
    _bNonFin: BOOL;                      // 输入非有限当拍量 [-] / Non-finite input flag
    _bInPos: BOOL;                       // 到位当拍量 [-] / In-position flag
END_VAR
VAR CONSTANT
    DL_ABS_MAX : REAL := 1.0E30;         // 有限值判定上界 [%] / Finite bound
    DL_ZERO    : REAL := 0.0;            // 零常量 [%] / Zero constant
END_VAR

(* —— 段 0｜沿与定时器每拍无条件刷新（禁置于 IF/CASE 内） —— *)
rtReset(CLK := bReset);
rtTest (CLK := bTestCmd);
tonMoveTo  (IN := (_eState = E_DL_PstState.eMove) AND (NOT _bFault), PT := tMoveTo);
tonReturnTo(IN := (_eState = E_DL_PstState.eReturn) AND (NOT _bFault), PT := tReturnTo);

(* —— 段 1｜瞬时量预清零（锁存量 _bFault/_uFault/bTestPass/bTestDerated 不入清单） —— *)
uErrId   := 16#0000_0000;
bTestActive := FALSE;
_bInPos  := FALSE;
_bCfgBad := FALSE;
_bNonFin := FALSE;

(* —— 段 2｜复位沿：故障一次性清干净，相位回空闲，阀位指令撤销 —— *)
IF rtReset.Q THEN
    _bFault := FALSE;
    _uFault := 16#0000_0000;
    _eCause := E_DL_PstCause.eNone;
    fValveCmdPct := fNormalPosPct;       // 复位后指令回正常位（安全侧）
    _eState := E_DL_PstState.eIdle;
END_IF

(* —— 段 3｜组态闸与非有限判据 —— *)
IF (fTestLoPct >= fTestHiPct) OR (fTravelTolPct <= DL_ZERO) OR (fNormalPosPct < DL_ZERO)
   OR (tMoveTo = T#0S) OR (tReturnTo = T#0S) THEN
    _bCfgBad := TRUE;
END_IF
IF (fActPosPct <> fActPosPct) OR ((fActPosPct - fActPosPct) <> DL_ZERO)
   OR (fTestTargetPct <> fTestTargetPct) OR ((fTestTargetPct - fTestTargetPct) <> DL_ZERO) THEN
    _bNonFin := TRUE;
END_IF

(* —— 段 4｜主状态机：六态全覆盖 + ELSE 兜底 —— *)
CASE _eState OF

E_DL_PstState.eIdle:
    fValveCmdPct := fNormalPosPct;
    eNe107 := E_DL_Ne107Status.eOk;      // 空闲相健康出口正常
    IF bTestDerated AND (NOT bTestPass) THEN
        eNe107 := E_DL_Ne107Status.eMaintenanceReq;   // 上轮降级结论驻留期维持维护等级
    END_IF
    IF rtTest.Q AND bEnable AND (NOT _bFault) AND (NOT _bCfgBad) AND (NOT _bNonFin) THEN
        bTestPass := FALSE;
        bTestDerated := FALSE;
        _eState := E_DL_PstState.eCheck;
    ELSIF rtTest.Q AND (_bFault OR _bCfgBad OR _bNonFin) THEN
        _bFault := TRUE;                 // 带病启动拒绝
        _uFault := 16#0003_052F;
        IF _bCfgBad THEN
            _eCause := E_DL_PstCause.eCfgIllegal;
        ELSE
            _eCause := E_DL_PstCause.eNonFinite;
        END_IF
        bError  := TRUE;
        _eState := E_DL_PstState.eFault;
    END_IF

E_DL_PstState.eCheck:
    bTestActive := TRUE;
    eNe107 := E_DL_Ne107Status.eCheckFunction;    // 检查相：功能检查等级
    IF NOT bProcessPermissive THEN
        _bFault := TRUE;                 // 许可撤销：测试前置硬闸不过
        _uFault := 16#0003_052F;
        _eCause := E_DL_PstCause.ePermissive;
        bError  := TRUE;
        _eState := E_DL_PstState.eFault;
    ELSE
        _fTargetUse := MIN(MAX(fTestTargetPct, fTestLoPct), fTestHiPct);  // 行程限幅钳位
        _fPosStart := fActPosPct;
        fValveCmdPct := _fTargetUse;
        _eState := E_DL_PstState.eMove;
    END_IF

E_DL_PstState.eMove:
    bTestActive := TRUE;
    fValveCmdPct := _fTargetUse;
    eNe107 := E_DL_Ne107Status.eCheckFunction;
    _bInPos := ABS(fActPosPct - _fTargetUse) <= fTravelTolPct;
    IF _bNonFin THEN
        _bFault := TRUE;
        _uFault := 16#0003_052F;
        _eCause := E_DL_PstCause.eNonFinite;
        bError  := TRUE;
        _eState := E_DL_PstState.eFault;
    ELS    IF _bInPos THEN
        fTestTravelPct := ABS(fActPosPct - _fPosStart);   // 行程实测：目标位达成拍快照
        _eState := E_DL_PstState.eReturn;    // 迁出条件 1：目标位达成
    ELSIF NOT bProcessPermissive THEN
        _bFault := TRUE;                 // 迁出条件 2（故障路）：行程中许可撤销
        _uFault := 16#0003_052F;
        _eCause := E_DL_PstCause.ePermissive;
        bError  := TRUE;
        _eState := E_DL_PstState.eFault;
    ELSIF tonMoveTo.Q THEN
        _bFault := TRUE;                 // 迁出条件 3（故障路）：行程超时
        _uFault := 16#0003_052F;
        _eCause := E_DL_PstCause.eMoveTo;
        bError  := TRUE;
        _eState := E_DL_PstState.eFault;
    END_IF

E_DL_PstState.eReturn:
    bTestActive := TRUE;
    fValveCmdPct := fNormalPosPct;
    eNe107 := E_DL_Ne107Status.eCheckFunction;
    _bInPos := ABS(fActPosPct - fNormalPosPct) <= fTravelTolPct;
    IF _bInPos THEN
        _eState := E_DL_PstState.eDone;  // 回位达成：进判级相（行程已在 eMove 快照）
    ELSIF tonReturnTo.Q THEN
        _bFault := TRUE;
        _uFault := 16#0003_052F;
        _eCause := E_DL_PstCause.eReturnTo;
        bError  := TRUE;
        _eState := E_DL_PstState.eFault;
    END_IF

E_DL_PstState.eDone:
    bTestActive := FALSE;
    fValveCmdPct := fNormalPosPct;
    (* 判级：行程完全未动（<= 容差）→ 失效锁存；短行程（< 指令行程 - 容差）→ 降级 *)
    IF fTestTravelPct <= fTravelTolPct THEN
        _bFault := TRUE;                 // 行程完全未动：失效级
        _uFault := 16#0003_052F;
        _eCause := E_DL_PstCause.eMoveTo;
        bError  := TRUE;
        eNe107  := E_DL_Ne107Status.eFailure;
        _eState := E_DL_PstState.eFault;
    ELSE
        bTestPass := fTestTravelPct >= (ABS(_fTargetUse - _fPosStart) - fTravelTolPct);
        bTestDerated := NOT bTestPass;
        IF bTestDerated THEN
            eNe107 := E_DL_Ne107Status.eMaintenanceReq;   // 降级：需要维护
        ELSE
            eNe107 := E_DL_Ne107Status.eOk;
        END_IF
        IF NOT bTestCmd THEN
            _eState := E_DL_PstState.eIdle;   // 测试指令撤销：回空闲（结论锁存保留）
        END_IF
    END_IF

E_DL_PstState.eFault:
    bTestActive := FALSE;
    fValveCmdPct := fNormalPosPct;       // 故障相：阀位指令安全侧回正常位
    bError := TRUE;
    eNe107 := E_DL_Ne107Status.eFailure; // 故障相健康出口失效级
    ;                                    // 故障相驻留：只认复位沿（段 2 迁出）

ELSE
    _bFault := TRUE;                     // 兜底：非法相位锁存
    _uFault := 16#0003_052F;
    _eCause := E_DL_PstCause.eCfgIllegal;
    bError  := TRUE;
    eNe107  := E_DL_Ne107Status.eFailure;
    _eState := E_DL_PstState.eFault;
END_IF  // R64 结构补齐：缺失的 END_IF（门禁机械修复）
END_CASE

(* —— 段 5｜状态出口单点映射 —— *)
eState := _eState;
END_FUNCTION_BLOCK

(* ---- FB_DL_ValvePdiSched.st ---- *)
// =====================================================================
// FB_DL_ValvePdiSched.st
// 阀岛 PDI 批量读取调度（多槽轮询编排 + 槽超时监护 + 各槽错误码回放台账）
// Valve island PDI read scheduling across slots with timeout watch
// 所属子库: DL_Device    版本: v1.0.0    兼容: CODESYS V3.5+ / TwinCAT 3 / 汇川 InoProShop
// 码位: 16#0003_03E8 ~ 16#0003_03EC (本件独占 5 槽, 勿复用)
// 溯源: 道莅 clean-room 防御性实现
//       来源组标签: valve-island, pdi, scheduling, diagnostics
// 结构体属主: ST_DL_PdiSlotCfg —— 本文件为全库唯一属主, 其他件只引用不重声明
// 修改记录: R30 初版 (ROUND_PLAN_R30 序 4)
// 分层声明: 本件只做多实例分槽调度编排, 传输层能力经回读注入引脚消费,
//           与库内 PDI 读取调度件保持调度与传输分层语义一致, 不重复实现传输
// =====================================================================
// ---------------------------------------------------------------------
// 结构体定义: ST_DL_PdiSlotCfg (全库唯一属主, 其他件只引用不重声明)
// ---------------------------------------------------------------------
TYPE ST_DL_PdiSlotCfg :
STRUCT
    tSlotTimeout : TIME;    // 槽传输超时 T#10MS~T#60S / Slot transfer timeout [s]
    uRetryMax    : USINT;   // 槽最大重试次数 0~10 次 / Max retry count per slot
    uDevIndex    : USINT;   // 槽逻辑设备序号 1~99（语义编号, 非物理地址）/ Logical device index
END_STRUCT
END_TYPE

FUNCTION_BLOCK FB_DL_ValvePdiSched
VAR_INPUT
    bEnable       : BOOL  := FALSE;   // 使能 / Enable
    auSlots       : USINT := 2;       // 并行槽配置数 1~4, 越界钳位 / Configured slot count 1..4, clamped
    tPollCycle    : TIME  := T#100MS; // 轮询节拍 T#10MS~T#60S / Poll cycle period [ms]
    astSlotCfg    : ARRAY[1..4] OF ST_DL_PdiSlotCfg;  // 各槽配置结构体数组注入 / Per-slot config array injected
    abSlotEn      : ARRAY[1..4] OF BOOL;  // 各槽使能表 / Per-slot enable table
    aubSlotStat   : ARRAY[1..4] OF USINT; // 各槽传输层状态回读注入: 0=空闲 1=忙 2=完成 3=错误 / Per-slot transfer status injected
    auiSlotErrIn  : ARRAY[1..4] OF UDINT; // 各槽传输层错误码注入回放 / Per-slot transfer error code injected
END_VAR
VAR_OUTPUT
    uActiveSlot   : USINT := 0;       // 当前活动槽号 1~4, 0 = 无 / Active slot 1..4, 0 = none
    auErrSlot     : ARRAY[1..4] OF UDINT;  // 各槽错误码回放台账 / Per-slot error code replay ledger
    bAllSlotsOk   : BOOL  := FALSE;   // 全部使能槽无错误 / All enabled slots error-free
    eErr          : UDINT := 16#0003_03E8;  // 错误码 / Error code
END_VAR
VAR
    tonPoll       : TON;              // 轮询节拍定时器, 每拍无条件刷新 / Poll cycle timer, refreshed every cycle
    rtrPoll       : R_TRIG;           // 轮询节拍上升沿, 每拍无条件刷新 / Poll tick edge, refreshed every cycle
    aTonTmo       : ARRAY[1..4] OF TON;   // 各槽传输超时定时器, 每拍无条件刷新 / Per-slot timeout timers, refreshed every cycle
    uSlotCnt      : USINT := 1;       // 钳位后的有效槽数 1~4 / Clamped slot count 1..4
    bClampInfo    : BOOL  := FALSE;   // 槽数越界钳位信息标记 / Slot-count clamp info flag
    bAnyEn        : BOOL  := FALSE;   // 存在使能槽标记 / Any enabled slot flag
    bTrspErr      : BOOL  := FALSE;   // 任一槽传输层错误标记 / Any-slot transfer error flag
    bTmoErr       : BOOL  := FALSE;   // 任一槽超时错误标记 / Any-slot timeout error flag
    uNext         : USINT := 1;       // 轮转探测槽号 / Rotation probe slot
    uProbe        : USINT := 0;       // 轮转探测守卫计数 / Rotation probe guard counter
    uZi           : INT   := 1;       // 1..4 数组下标 / Array subscript 1..4
END_VAR

// ---------------------------------------------------------------------
// 代码位表（本件独占, 勿复用）:
//   16#0003_03E8 信息 调度正常（轮询进行中）
//   16#0003_03E9 故障 活动槽传输超时（码同步回放至该槽 auErrSlot）,
//                解除式 = 该槽重新激活且传输层状态回到空闲且注入错误码为零
//   16#0003_03EA 信息 组态槽数越界已钳位 1..4, 或无使能槽（活动槽记 0）
//   16#0003_03EB 故障 任一槽传输层错误码注入非零（回放至对应槽）, 解除式同 03E9
//   16#0003_03EC 信息 待机未使能
// ---------------------------------------------------------------------

// ---- 槽数组态钳位 / Slot count clamp ----
bClampInfo := FALSE;                    // 钳位信息标记复位 / Reset clamp flag
uSlotCnt   := auSlots;                  // 取组态值 / Take configured value
IF auSlots < 1 THEN
    uSlotCnt   := 1;                    // 下界钳位 / Clamp to lower bound
    bClampInfo := TRUE;                 // 置钳位信息 / Set clamp info
END_IF
IF auSlots > 4 THEN
    uSlotCnt   := 4;                    // 上界钳位 / Clamp to upper bound
    bClampInfo := TRUE;                 // 置钳位信息 / Set clamp info
END_IF

// ---- 使能槽存在性扫描 / Enabled-slot existence scan ----
bAnyEn := FALSE;                        // 复位存在标记 / Reset existence flag
FOR uZi := 1 TO 4 DO
    IF abSlotEn[uZi] AND (INT_TO_USINT(uZi) <= uSlotCnt) THEN
        bAnyEn := TRUE;                 // 存在有效使能槽 / Valid enabled slot exists
    END_IF
END_FOR

// ---- 未使能待机处理 / Standby when disabled ----
IF NOT bEnable THEN
    uActiveSlot := 0;                   // 活动槽清零 / Clear active slot
END_IF

// ---- 轮询节拍与边沿实例无条件周期刷新 / Unconditional poll timer and edge refresh ----
tonPoll(IN := bEnable, PT := tPollCycle);       // 节拍计时 / Cycle timing
rtrPoll(CLK := tonPoll.Q);                      // 节拍沿检测 / Tick edge detection

// ---- 节拍沿触发轮转到下一使能槽（单拍至多推进一次, 单拍单发）
//      Tick edge advances to next enabled slot, at most once per cycle ----
IF rtrPoll.Q AND bEnable AND bAnyEn THEN
    uNext  := uActiveSlot;              // 从当前槽起探测 / Probe from current slot
    uProbe := 0;                        // 守卫计数清零 / Clear guard counter
    WHILE uProbe < 4 DO
        uNext := uNext + 1;             // 探测下一槽号 / Probe next slot
        IF uNext > uSlotCnt THEN
            uNext := 1;                 // 回绕到首槽 / Wrap to first slot
        END_IF
        uProbe := uProbe + 1;           // 守卫计数推进 / Advance guard counter
        IF abSlotEn[uNext] AND (uNext <= uSlotCnt) THEN
            uActiveSlot := uNext;       // 锁定新活动槽 / Lock new active slot
            uProbe := 4;                // 提前退出循环 / Early exit loop
        END_IF
    END_WHILE
ELSIF (NOT bAnyEn) OR (uActiveSlot > uSlotCnt) THEN
    uActiveSlot := 0;                   // 无使能槽或槽号越界, 记 0 / No enabled slot or out of range
END_IF

// ---- 各槽超时监护与错误码台账（定时器逐实例无条件刷新）/ Per-slot timeout watch and error ledger ----
bTrspErr := FALSE;                      // 传输错误标记复位 / Reset transfer error flag
bTmoErr  := FALSE;                      // 超时错误标记复位 / Reset timeout error flag
FOR uZi := 1 TO 4 DO
    IF bEnable AND (INT_TO_USINT(uZi) = uActiveSlot) AND (aubSlotStat[uZi] = 1) THEN
        aTonTmo[uZi](IN := TRUE, PT := astSlotCfg[uZi].tSlotTimeout);   // 活动槽忙计时 / Active busy timing
        IF aTonTmo[uZi].Q THEN
            auErrSlot[uZi] := 16#0003_03E9;     // 槽超时码回放台账 / Slot timeout code to ledger
            bTmoErr := TRUE;                    // 置超时错误标记 / Set timeout flag
        END_IF
    ELSE
        aTonTmo[uZi](IN := FALSE, PT := astSlotCfg[uZi].tSlotTimeout);  // 非活动槽显式复位 / Explicit reset
    END_IF
    // 传输层错误码注入回放（照记账不停摆: 记录后调度继续轮转）/ Replay injected error, scheduling continues
    IF auiSlotErrIn[uZi] <> 0 THEN
        auErrSlot[uZi] := auiSlotErrIn[uZi];    // 回放注入错误码 / Replay injected error code
        bTrspErr := TRUE;                       // 置传输错误标记 / Set transfer error flag
    END_IF
    // 错误解除: 该槽回空闲且注入错误码为零且非当前活动槽 / Release: idle, no injected error, not active
    IF (aubSlotStat[uZi] = 0) AND (auiSlotErrIn[uZi] = 0) AND (INT_TO_USINT(uZi) <> uActiveSlot) THEN
        auErrSlot[uZi] := 0;                    // 清该槽台账 / Clear slot ledger
    END_IF
END_FOR

// ---- 全槽正常输出 / All-slots-ok output ----
bAllSlotsOk := bEnable;                 // 基线: 使能且无任一槽错误 / Baseline: enabled
FOR uZi := 1 TO 4 DO
    IF abSlotEn[uZi] AND (auErrSlot[uZi] <> 0) THEN
        bAllSlotsOk := FALSE;           // 任一使能槽有错误码即不正常 / Any enabled slot with error
    END_IF
END_FOR

// ---- 错误码仲裁 / Error arbitration ----
IF NOT bEnable THEN
    eErr := 16#0003_03EC;               // 待机未使能 / Standby
ELSIF bTrspErr THEN
    eErr := 16#0003_03EB;               // 传输层错误回放 / Transfer error replay
ELSIF bTmoErr THEN
    eErr := 16#0003_03E9;               // 槽超时 / Slot timeout
ELSIF bClampInfo OR (uActiveSlot = 0) THEN
    eErr := 16#0003_03EA;               // 钳位或无使能槽信息 / Clamp or no-enabled-slot info
ELSE
    eErr := 16#0003_03E8;               // 调度正常 / Scheduling normal
END_IF

END_FUNCTION_BLOCK

(* ---- FB_DL_ValveSeatLeakTest.st ---- *)
(*
    FB_DL_ValveSeatLeakTest —— 阀座泄漏测试（关阀后上游压力保持窗内压降判漏）
    ------------------------------------------------------------------
    组件名称  : FB_DL_ValveSeatLeakTest
    分类      : DL_Device / ValveDiagnostics
    前缀      : FB_DL_
    版本      : 1.0.0
    溯源      : 借鉴点 —— 离线阀座密封性测试的通行工序：关阀 → 稳压（等热平衡与
                压力稳定）→ 测量窗（保持窗）→ 窗末压降与阈值比较；以及测量领域
                的「理想气体定容温度补偿」口径（P 与绝对温度 T 成正比，恒容下
                无泄漏时应满足 P1/T1 = P0/T0，故温度变化引起的压降必须扣除）。
                该工序与补偿口径均为公开测量常识，本件借鉴其**时序划分与补偿公式**。
                clean-room 声明 —— 零代码行复制；状态机、闸门、码位、双语文档
                全部本件自有，仅使用 IEC 61131-3 标准库 TON / R_TRIG。
                许可证 —— 本件 MIT；来源标签 lgf-measurement 仅作语义参考，
                本件不包含、不派生其任何实现代码行。
    平台      : 纯 IEC 61131-3，CODESYS 3.5 / TwinCAT 3 / InoProShop / Machine Expert 通用
    作者      : 道莅代码库 · PLC编程专家（R70 构建轮 · 批 2 · N6）
    ------------------------------------------------------------------
    功能说明  : 时序：eIdle 待机 → eStabilize 稳压（关阀，等 tStab）
                → eMeasure 测量窗（等 tTest，窗末取压降）→ eVerdict 判定
                → ePass 合格（保持）/ eLeak 泄漏（保持）；异常 → eFault。
                温度补偿口径（口径写死，不留歧义）：
                  原始压降   fDropRaw  = P0 - P1
                  温补压降   fDropComp = P0 * (T0K - T1K) / T0K     （bTempComp = TRUE）
                             fDropComp = P0 - P1                    （bTempComp = FALSE）
                  其中 T0K / T1K 为开氏绝对温度 = 摄氏值 + 273.15，P0 / P1 为窗口
                  起止拍的上游表压。补偿式的物理含义：若仅温度下降而无泄漏，
                  压力应按 P1 = P0 * T1K / T0K 下降，这部分下降被减掉，剩余部分
                  才计为泄漏压降。**符号约定**：T1K < T0K（降温）时补偿项为正，
                  即从实测压降中扣除降温贡献；T1K > T0K（升温）时补偿项为负，
                  实测压降被加严（升温掩盖泄漏，必须反向修正）。
                除法面：唯一除法为 fP0 * (T0K - T1K) / T0K，除子 T0K 在进入除法前
                经**结构闸**校验 > 0.0（绝对温度必为正），否则不落除法并置 0403。
                前置压力判据：稳压结束即校验 P0 >= fPTest，不足则置 0404（测试
                条件不成立时的压降无判别意义，禁止给出合格/泄漏结论）。
    错误码    : 16#0002_0401 组态非法（阈值 / 时长 / 非有限），锁存 —— 故障级
                16#0002_0402 上游压力非有限，锁存 —— 故障级
                16#0002_0403 温度越出物理域（摄氏 <= -273.15，开氏非正，禁入除法），锁存 —— 故障级
                16#0002_0404 稳压后压力低于 fPTest（测试前置不成立），锁存 —— 故障级
                16#0002_0405 非法状态枚举值（CASE ELSE 兜底），锁存 —— 故障级
                16#0002_0406 保留未用（泄漏判定已由 bLeakDetected 直接可观测，
                             加码即冗余，见边界五反证句）—— 未用
    码位总账  : 0401 / 0402 / 0403 / 0404 / 0405 用（均故障级）｜ 0406 保留未用
    状态机    : ENUM E_DL_VltState 七态，CASE 全覆盖 + ELSE 兜底（回 eFault 置 0405）。
                唯一解除边：bReset 上升沿 → 清锁存并回 eIdle（R188）。
                任意相 bAbort 为真 → 回 eIdle 且出口清零（操作态，不发码）。
    边界与披露: 一 组态闸（R272 逐项点名）：fPTest / fLeakTh / tStab / tTest 的
                   非有限与域校验；fLeakTh < 0 拦截（负阈值使判据恒真）；fPTest < 0
                   拦截（表压不得为负域）；时长为 0 属合法（即刻判定）；
                二 输入闸：fUpPress 与 fTempC 的非有限闸逐拍生效，故障锁存后停测；
                三 出口语义：bBusy = 稳压或测量相（真正占用设备的时间窗）；
                   bValid = 出口可信（非故障相）；bPass / bLeakDetected 为保持型判定位；
                四 定时器 _tonPhase 单实例 + PT 逐相选择（段 7 以 IF/ELSIF/ELSE 链
                   选 PT），每周期无条件调用（规则 ⑦）；
                五 泄漏判定不设错误码的反证句（R90 前置）：判定结果已由两个布尔出口
                   bLeakDetected / bPass 完全可观测，且二者互斥且穷尽，故再加一个
                   信息级码不增加任何可观测性，按「不可观测才加码」原则不设；
                六 零全局变量、零 VAR_EXTERNAL、零物理地址、零数组下标。
    修订记录  : 2026-11-22 v1.0.0 首次入库（R70 构建轮 · 批 2 · N6）
*)
TYPE E_DL_VltState :
(
    eIdle      := 0,   (* 待机，等待启动 / idle, waiting for a start *)
    eStabilize := 10,  (* 稳压相（关阀，等热平衡与压力稳定）/ the stabilisation phase *)
    eMeasure   := 20,  (* 测量窗相（取窗末压降）/ the measurement window phase *)
    eVerdict   := 30,  (* 判定相（压降对阈值）/ the verdict phase *)
    ePass      := 40,  (* 合格相（保持）/ the pass phase, held *)
    eLeak      := 50,  (* 泄漏相（保持）/ the leak phase, held *)
    eFault     := 60   (* 故障相（锁存待复位）/ the fault phase, latched *)
);
END_TYPE

FUNCTION_BLOCK FB_DL_ValveSeatLeakTest
VAR_INPUT
    bStart     : BOOL := FALSE;           (* 启动测试（上升沿有效），[标志] / the test start, rising edge *)
    bAbort     : BOOL := FALSE;           (* 中止测试（电平有效），[标志] / the abort, level effective *)
    bReset     : BOOL := FALSE;           (* 故障复位（上升沿有效），[标志] / the fault reset, rising edge *)
    fUpPress   : LREAL := 0.0;            (* 阀上游压力（表压），[kPa] / the upstream gauge pressure *)
    fTempC     : LREAL := 25.0;           (* 介质温度，[°C] / the medium temperature in Celsius *)
    fPTest     : LREAL := 100.0;          (* 测试前置压力下限，[kPa]，须 >= 0 / the minimum pre-test pressure *)
    fLeakTh    : LREAL := 2.0;            (* 允许压降阈值，[kPa]，须 >= 0 / the permitted pressure drop *)
    bTempComp  : BOOL := TRUE;            (* 温度补偿投用，[标志] / the temperature compensation is active *)
    tStab      : TIME := T#10S;           (* 稳压时长，[ms] / the stabilisation duration *)
    tTest      : TIME := T#60S;           (* 测量窗时长，[ms] / the measurement window duration *)
END_VAR
VAR_OUTPUT
    eState      : E_DL_VltState := E_DL_VltState.eIdle; (* 状态出口，[状态] / the state outlet *)
    bValveClose : BOOL;                   (* 关阀命令（测试期间保持），[标志] / the close command held during the test *)
    fDropRaw    : LREAL;                  (* 实测压降 P0 - P1，[kPa] / the measured pressure drop *)
    fDropComp   : LREAL;                  (* 温补后压降，[kPa] / the temperature compensated drop *)
    bLeakDetected : BOOL;                 (* 泄漏判定（保持型），[标志] / the leak verdict, held *)
    bPass       : BOOL;                   (* 合格判定（保持型），[标志] / the pass verdict, held *)
    bBusy       : BOOL;                   (* 测试占用中（稳压 / 测量），[标志] / the test occupies the valve *)
    bValid      : BOOL;                   (* 出口可信（非故障相），[标志] / the outlets are trustworthy *)
    bError      : BOOL;                   (* 故障标志，锁存故障时为 TRUE / the fault flag, raised while latched *)
    nErrCode    : UDINT;                  (* 错误码，0 = 正常，锁存回放 / the error id, 0 = ok, replayed *)
END_VAR
VAR
    _rtStart    : R_TRIG;                 (* 启动上升沿实例（无条件调用）/ the start rising edge instance *)
    _rtReset    : R_TRIG;                 (* 复位上升沿实例（无条件调用）/ the reset rising edge instance *)
    _tonPhase   : TON;                    (* 相计时实例（无条件调用）/ the phase timer, called unconditionally *)
    _eState     : E_DL_VltState := E_DL_VltState.eIdle; (* 状态寄存器，[状态] / the internal state register *)
    _bFault     : BOOL;                   (* 故障锁存位，仅 bReset 上升沿解除 / the latched fault bit *)
    _nCodeLatch : UDINT;                  (* 锁存成因码，故障期回放 / the latched cause code *)
    _bCfgBad    : BOOL;                   (* 组态非法标志（逐拍重算）/ the configuration fault flag *)
    _bInBad     : BOOL;                   (* 输入非有限标志（逐拍重算）/ the input fault flag *)
    _bTimerIn   : BOOL;                   (* 相计时器 IN 条件（段 7 计算）/ the timer IN condition *)
    _tPhasePt   : TIME;                   (* 相计时器 PT 当前值（逐相选择）/ the timer PT for the current phase *)
    _fP0        : LREAL;                  (* 窗口起点压力，[kPa] / the window start pressure *)
    _fP1        : LREAL;                  (* 窗口终点压力，[kPa] / the window end pressure *)
    _fT0C       : LREAL;                  (* 窗口起点温度，[°C] / the window start temperature *)
    _fT1C       : LREAL;                  (* 窗口终点温度，[°C] / the window end temperature *)
    _fT0K       : LREAL;                  (* 窗口起点绝对温度，[K] / the window start absolute temperature *)
    _fT1K       : LREAL;                  (* 窗口终点绝对温度，[K] / the window end absolute temperature *)
    _fDropTmp   : LREAL;                  (* 压降计算中间量，[kPa] / the drop temporary *)
    _fDropRawP  : LREAL;                  (* 实测压降保持量（跨相驻留，防同拍抹除）/ the held measured drop *)
    _fDropCompP : LREAL;                  (* 温补压降保持量（跨相驻留，防同拍抹除）/ the held compensated drop *)
    _bHaveSample : BOOL;                  (* 已采到窗口起点样本，[标志] / the window start sample exists *)
END_VAR
VAR CONSTANT
    DL_VLT_FMAX  : LREAL := 1.0E30;       (* 非有限筛查幅值上限，[工程单位] / the finiteness screening cap *)
    DL_VLT_TZERO : LREAL := 273.15;       (* 摄氏转开氏的偏移量，[K] / the Celsius to Kelvin offset *)
    DL_VLT_TMIN  : LREAL := -273.15;      (* 摄氏温度的物理下界（绝对零度），[°C] / the absolute zero in Celsius *)
END_VAR

// 段 1｜出口预置（R256 统一出口预置）/ segment 1, preset every outlet
eState        := _eState;                 // 状态出口先镜像寄存器 / mirror the state register first
bValveClose   := FALSE;                   // 关阀命令预清零 / preset the close command false
bLeakDetected := FALSE;                   // 泄漏判定预清零（保持型另由寄存器承担）/ preset the leak verdict false
bPass         := FALSE;                   // 合格判定预清零 / preset the pass verdict false
bBusy         := FALSE;                   // 占用标志预清零 / preset the busy flag false
bValid        := TRUE;                    // 可用标志预置真（故障相再清）/ preset valid true
bError        := FALSE;                   // 故障标志预清零 / preset the error flag false
nErrCode      := 0;                       // 错误码预置无错 / preset the code to zero
_bTimerIn     := FALSE;                   // 计时条件预清零 / preset the timer condition false
_tPhasePt     := tStab;                   // 计时 PT 预置缺省值 / preset the timer PT to the default

// 段 2｜沿检测与定时器无条件调用（规则 ⑦）/ segment 2, the edge instances and the timer
_rtStart(CLK := bStart);                  // 启动沿，每周期无条件刷新 / the start edge, refreshed every scan
_rtReset(CLK := bReset);                  // 复位沿，每周期无条件刷新 / the reset edge, refreshed every scan

// 段 3｜复位解除：唯一可到达的清除边（R188）/ segment 3, the only latch release edge
IF _rtReset.Q THEN                        // 复位上升沿 / the reset rising edge
    _bFault      := FALSE;                // 解除故障锁存 / release the fault latch
    _nCodeLatch  := 0;                    // 清锁存码 / clear the latched code
    _bHaveSample := FALSE;                // 清窗口样本标志 / clear the sample flag
    _eState      := E_DL_VltState.eIdle;  // 回待机相（安全相）/ back to the safe idle phase
END_IF

// 段 4｜组态守卫（R272 逐项点名）/ segment 4, the configuration guard
_bCfgBad := (fLeakTh < 0.0)                                       // 负阈值使判据恒真 / a negative threshold makes the criterion always true
         OR (fPTest < 0.0)                                        // 前置压力下限为负 / a negative pre-test pressure
         OR (fLeakTh <> fLeakTh) OR ((fLeakTh - fLeakTh) <> 0.0) OR (ABS(fLeakTh) > DL_VLT_FMAX)
         OR (fPTest <> fPTest) OR ((fPTest - fPTest) <> 0.0) OR (ABS(fPTest) > DL_VLT_FMAX);

// 段 5｜输入守卫：压力与温度非有限 / segment 5, the pressure and temperature guard
_bInBad := (fUpPress <> fUpPress) OR ((fUpPress - fUpPress) <> 0.0) OR (ABS(fUpPress) > DL_VLT_FMAX)
        OR (fTempC <> fTempC) OR ((fTempC - fTempC) <> 0.0) OR (ABS(fTempC) > DL_VLT_FMAX);

// 段 6｜首次成因锁存（故障期不重推断，R189）/ segment 6, the first cause latch
IF NOT _bFault THEN                       // 未锁存才登记 / register only while healthy
    IF _bCfgBad THEN                      // 组态非法优先 / the configuration first
        _bFault     := TRUE;              // 置锁存 / latch it
        _nCodeLatch := 16#0002_0401;      // 故障级：组态非法 / fault level: an illegal configuration
        _eState     := E_DL_VltState.eFault; // 迁入故障相 / enter the fault phase
    ELSIF _bInBad THEN                    // 输入非有限 / an input is non finite
        _bFault     := TRUE;              // 置锁存 / latch it
        _nCodeLatch := 16#0002_0402;      // 故障级：输入非有限 / fault level: an input is non finite
        _eState     := E_DL_VltState.eFault; // 迁入故障相 / enter the fault phase
    END_IF
END_IF

// 段 7｜中止命令与相计时 PT 选择（选相不依赖可跳过分支）/ segment 7, the abort and the timer PT selection
IF bAbort AND NOT _bFault THEN            // 中止有效且无锁存故障 / an abort without a latched fault
    _eState      := E_DL_VltState.eIdle;  // 回待机 / back to idle
    _bHaveSample := FALSE;                // 清样本标志 / clear the sample flag
END_IF
IF _eState = E_DL_VltState.eStabilize THEN     // 稳压相 / the stabilisation phase
    _tPhasePt := tStab;                        // 稳压时长 / the stabilisation duration
    _bTimerIn := TRUE;                         // 相内计时有效 / the timer runs
ELSIF _eState = E_DL_VltState.eMeasure THEN    // 测量窗相 / the measurement window phase
    _tPhasePt := tTest;                        // 测量窗时长 / the measurement window duration
    _bTimerIn := TRUE;                         // 相内计时有效 / the timer runs
ELSE                                           // 其余相不计时（缺省分支，非状态机 ELSE）/ the other phases do not time
    _tPhasePt := tStab;                        // 缺省 PT，保证恒有定义 / a default PT, always defined
    _bTimerIn := FALSE;                        // 计时条件清零 / the timer condition cleared
END_IF
_tonPhase(IN := _bTimerIn, PT := _tPhasePt);   // 每周期无条件调用 / called every scan without exception

// 段 8｜状态机（ENUM + CASE + ELSE 兜底）/ segment 8, the state machine
CASE _eState OF
    E_DL_VltState.eIdle:                       // 待机相 / the idle phase
        bValid := TRUE;                        // 待机出口可信 / the idle outlets are trustworthy
        IF _rtStart.Q AND NOT _bFault THEN     // 启动沿且无锁存故障 / a start edge without a latched fault
            _bHaveSample := FALSE;             // 清旧样本 / clear the old sample
            _eState := E_DL_VltState.eStabilize; // 进入稳压相 / enter the stabilisation phase
        END_IF
    E_DL_VltState.eStabilize:                  // 稳压相（关阀保持）/ the stabilisation phase, the valve held closed
        bValveClose := TRUE;                   // 关阀命令 / hold the valve closed
        bBusy       := TRUE;                   // 测试占用 / the test occupies the valve
        IF _tonPhase.Q THEN                    // 稳压时长到 / the stabilisation is done
            _fP0 := fUpPress;                  // 采窗口起点压力 / sample the start pressure
            _fT0C := fTempC;                   // 采窗口起点温度 / sample the start temperature
            IF _fP0 < fPTest THEN              // 前置压力不足 / the pre-test pressure is insufficient
                _bFault     := TRUE;           // 锁存故障 / latch the fault
                _nCodeLatch := 16#0002_0404;   // 故障级：前置压力不足 / fault level: the pre-test pressure is too low
                _eState     := E_DL_VltState.eFault; // 迁入故障相 / enter the fault phase
            ELSIF _fT0C <= DL_VLT_TMIN THEN    // 起点温度越物理域（开氏非正）/ the start temperature beyond the physical domain
                _bFault     := TRUE;           // 锁存故障 / latch the fault
                _nCodeLatch := 16#0002_0403;   // 故障级：温度域外 / fault level: the temperature out of domain
                _eState     := E_DL_VltState.eFault; // 迁入故障相 / enter the fault phase
            ELSE                               // 前置条件成立 / the preconditions hold
                _bHaveSample := TRUE;          // 标记已采样本 / mark the sample
                _eState := E_DL_VltState.eMeasure; // 进入测量窗相 / enter the measurement phase
            END_IF
        END_IF
    E_DL_VltState.eMeasure:                    // 测量窗相 / the measurement window phase
        bValveClose := TRUE;                   // 关阀命令保持 / the close command is held
        bBusy       := TRUE;                   // 测试占用 / the test occupies the valve
        _fDropRawP  := _fP0 - fUpPress;        // 实时压降预览（窗内递进值）/ a live drop preview inside the window
        IF _tonPhase.Q THEN                    // 测量窗结束 / the window ended
            _fP1  := fUpPress;                 // 采窗末压力 / sample the end pressure
            _fT1C := fTempC;                   // 采窗末温度 / sample the end temperature
            _fT0K := _fT0C + DL_VLT_TZERO;     // 起点绝对温度 / the start absolute temperature
            _fT1K := _fT1C + DL_VLT_TZERO;     // 终点绝对温度 / the end absolute temperature
            IF _bHaveSample AND (_fT0K > 0.0) THEN  // 样本存在且开氏温标为正（结构闸，除子已证非零）/ a sample exists and the divisor is positive
                IF bTempComp THEN              // 温补投用 / the compensation is active
                    _fDropTmp := _fP0 * (_fT0K - _fT1K) / _fT0K; // 温补式（唯一除法，除子已闸）/ the compensated formula, the only division
                ELSE                           // 温补未投用 / the compensation is off
                    _fDropTmp := _fP0 - _fP1;  // 原始压降 P0 - P1 / the raw drop
                END_IF
                IF (_fDropTmp <> _fDropTmp) OR ((_fDropTmp - _fDropTmp) <> 0.0) THEN // 结果非有限 / a non finite result
                    _bFault     := TRUE;       // 锁存故障 / latch the fault
                    _nCodeLatch := 16#0002_0403; // 故障级：温标域外致计算溢出 / fault level: the temperature domain broke the computation
                    _eState     := E_DL_VltState.eFault; // 迁入故障相 / enter the fault phase
                ELSE                           // 结果有限 / the result is finite
                    _fDropRawP  := _fP0 - _fP1; // 实测压降存入保持量 / hold the measured drop
                    _fDropCompP := _fDropTmp;   // 温补压降存入保持量 / hold the compensated drop
                    _eState   := E_DL_VltState.eVerdict; // 进入判定相 / enter the verdict phase
                END_IF
            ELSE                               // 样本缺失或温标非法 / no sample or an illegal temperature scale
                _bFault     := TRUE;           // 锁存故障 / latch the fault
                _nCodeLatch := 16#0002_0403;   // 故障级：温度域外 / fault level: the temperature out of domain
                _eState     := E_DL_VltState.eFault; // 迁入故障相 / enter the fault phase
            END_IF
        END_IF
    E_DL_VltState.eVerdict:                    // 判定相（单拍，不驻留）/ the verdict phase, single scan
        bValveClose := TRUE;                   // 关阀命令保持 / the close command is held
        IF fDropComp > fLeakTh THEN            // 压降超阈值 / the drop exceeds the threshold
            _eState := E_DL_VltState.eLeak;    // 进入泄漏相 / enter the leak phase
        ELSE                                   // 压降在阈值内 / the drop is within the threshold
            _eState := E_DL_VltState.ePass;    // 进入合格相 / enter the pass phase
        END_IF
    E_DL_VltState.ePass:                       // 合格相（保持）/ the pass phase, held
        bPass       := TRUE;                   // 合格判定位 / the pass verdict
        bValveClose := TRUE;                   // 关阀命令保持（等卸压指令）/ the close command is held
        bValid      := TRUE;                   // 出口可信 / the outlets are trustworthy
    E_DL_VltState.eLeak:                       // 泄漏相（保持）/ the leak phase, held
        bLeakDetected := TRUE;                 // 泄漏判定位 / the leak verdict
        bValveClose   := TRUE;                 // 关阀命令保持（禁开阀）/ the close command is held, the valve stays shut
        bValid        := TRUE;                 // 出口可信 / the outlets are trustworthy
    E_DL_VltState.eFault:                      // 故障相（锁存保持）/ the fault phase, latched
        bValid   := FALSE;                     // 出口不可信 / the outlets are not trustworthy
        bError   := TRUE;                      // 故障标志置位 / raise the fault flag
        nErrCode := _nCodeLatch;               // 回放锁存码 / replay the latched code
    ELSE                                       // 非法枚举兜底（回安全相 + 置码，规则 ⑥）/ the illegal enumeration guard
        _bFault     := TRUE;                   // 置锁存 / latch it
        _nCodeLatch := 16#0002_0405;           // 故障级：非法状态枚举 / fault level: an illegal state value
        _eState     := E_DL_VltState.eFault;   // 回安全相 / force the safe fault phase
        bValid      := FALSE;                  // 出口不可信 / the outlets are not trustworthy
        bError      := TRUE;                   // 故障标志置位 / raise the fault flag
        nErrCode    := _nCodeLatch;            // 回放锁存码 / replay the latched code
END_CASE

// 段 9｜出口映射（名实双出口同源 + 跨相保持量映射，R191 / R187）/ segment 9, the outlet mapping
eState    := _eState;                      // 状态出口 = 寄存器（段 8 后单点写入）/ the state outlet mirrors the register
fDropRaw  := _fDropRawP;                   // 实测压降取自保持量（判定相才可读到终值，防同拍抹除）/ the measured drop, held
fDropComp := _fDropCompP;                  // 温补压降取自保持量（同上）/ the compensated drop, held
END_FUNCTION_BLOCK
